(* CODESYS project Servo_Test.project

Project tree, tasks and I/O mapping:
  Device : CODESYS Virtual Control for Linux SL, CODESYS, order no. 2302000005, version 4.22.0.0
    application Application
      libraries: Standard, 3.5.22.0 (System); VisuDialogs, * (System); Unit Conversion Interfaces, * (Intern); CAA Mathematics, * (CAA Technical Workgroup); SM3_Math, * (CODESYS); SysProcess, * (System); CmpBitmapPool, * (System); SysProcess Implementation, * (System)
      task MainTask (cyclic, interval t#20ms, priority 1) calls MAIN_PRG, Ablaufkette
      task SoftMotion_PlanningTask (cyclic, interval t#2ms, priority 15) calls nothing
      global variables GVL_OPCUA
      visualisation Topics_Vis
      Structs/
        ST_RobotStatus/
          data type ST_RobotStatus
        ST_RobotAction/
          data type ST_RobotAction
          data type Error_Codes_RobotAction
        ST_RobotCommand/
          data type ST_RobotCommand
          data type Status_Codes_RobotCommand
        ST_Orientierung/
          data type ST_euler
          data type ST_quaternions
        ST_Roboter/
          data type ST_Pose_Axis
          data type ST_Pose_TCP
      old_code/
        data type Manuell_Achse
        data type TCP_Pose
        program PRG_VISU [ST]
        data type JointState
        data type ST_Servo_Axis
        data type ST_Servo_TCP
        FB_Robot/
          function block FB_Robot [FBD]
          function block FB_Watchdog [ST]
          function block FB_RobotCommander [ST]
        Interfaces/
          interface IF_RobotStatus: Ist_Pose_Axis, Ist_Pose_TCP, Ist_Mode, Client_Connection_Status, Update_Watchdog
          interface IF_RobotCommand: Soll_Pose_Axis, Soll_Pose_TCP
        function block FB_Roboter [FBD]: Update_Watchdog, Soll_Pose_Axis, Soll_Pose_TCP, Client_Connection_Status, Ist_Mode, Ist_Pose_Axis, Ist_Pose_TCP
        function block Status_POU [ST]
      program MAIN_PRG [FBD]
      FB_Generell/
        function block FB_MoveAction [ST]: MoveToHome, Ex1_ompl_tcp, Ex2_ompl_joint, Ex3_pilz_tcp_ptp, Ex_4_pilz_tcp_lin, Ablauf_HomePos, Ablauf_Pos1, Ablauf_Pos2, Ablauf_Pos3, Ablauf_Pos4, Ablauf_Pos5
        function block FB_Modes [FBD]
        function block FB_RobotStatus [ST]
        function block FB_RobotCommand [ST]
      program Ablaufkette [SFC]: Pos_6
      Funktionen/
        function FUNC_quat_to_euler [ST]
        function block FB_Quat_to_ZYZ [FBD]
        function block FB_ZYZ_to_Quat [FBD]
      Symbols
      image pool ImagePool
      visualisation VISU_Auto
      visualisation VISU_Startseite
      visualisation VISU_Manuell
      visualisation VISU_Konfig
      visualisation VISU_Schrittkette
  libraries: SM3_Robotics, * (CODESYS); VisuSymbols, 4.5.0.0 (System)
  text list GlobalTextList
*)

// Device/Application/old_code/Manuell_Achse
TYPE Manuell_Achse :
STRUCT
	axis_0_plus : BOOL;
	axis_0_minus : BOOL;
	axis_1_plus : BOOL;
	axis_1_minus : BOOL;
	axis_2_plus : BOOL;
	axis_2_minus : BOOL;
	axis_3_plus : BOOL;
	axis_3_minus : BOOL;
	axis_4_plus : BOOL;
	axis_4_minus : BOOL;
	axis_5_plus : BOOL;
	axis_5_minus : BOOL;
	//velocity_spee  einstellen
	//start manuell
END_STRUCT
END_TYPE

// Device/Application/old_code/TCP_Pose
TYPE TCP_Pose :
STRUCT
	trans_x : LREAL;
	trans_y : LREAL;
	trans_z : LREAL;
	rot_x : LREAL;
	rot_y : LREAL;
	rot_z : LREAL;
	rot_w : LREAL;
END_STRUCT
END_TYPE

//TCP Pose in kartesischen Koordinaten
//Rotation wird in quaternions uebermittelt, muss noch umgerechnet werden

// Device/Application/old_code/JointState
TYPE JointState :
STRUCT
	name :ARRAY[0..5] OF STRING;
	position :ARRAY[0..5] OF LREAL; 
	effort :ARRAY[0..5] OF LREAL;
	velocity :ARRAY[0..5] OF LREAL;
END_STRUCT
END_TYPE

// Device/Application/Structs/ST_RobotStatus/ST_RobotStatus
// Gibt den aktuellen Status des Roboters an
TYPE ST_RobotStatus :
STRUCT
	//Joints
	Ist_Pos_Axis : ST_Pose_Axis; 	
	
	// TCP mit Orientierung in Quaternions
	Ist_Pos_TCP : ST_Pose_TCP;	
	
	//Watchdog
	client_connected : BOOL;
	watchdog_counter : INT;		// Überprüft serverseitige client verbindung
END_STRUCT
END_TYPE

// Device/Application/Structs/ST_RobotCommand/ST_RobotCommand
TYPE ST_RobotCommand :
STRUCT
	// Achsen manuell verfahren
	Mode_Axis: BOOL;
	Soll_Axis_Servo : ST_Pose_Axis;
	Soll_Axis_Velocity: LREAL;
	
	// TCP manuell verfahren (funktioniert nicht, da Singularitäten auftreten wenn MoveIt Servo verwendet! Nicht in Code implementiert!)
	Mode_TCP: BOOL;
	Soll_TCP_Servo : ST_Pose_TCP;	// Hinweis: Rotation wird nur mit x,y,z übergeben und nicht als Quaternion!
	Soll_TCP_Velocity: LREAL;
	
	//enable: zum starten und stopen des services servo_node/start_servo und stop_servo
	enable : BOOL;
	
	//Status Code mit Status Codes
	Status_Code: SINT;
	
	//Watchdog
	client_connected: BOOL;
	watchdog_counter: INT;
END_STRUCT
END_TYPE

// Device/Application/Structs/ST_RobotAction/ST_RobotAction
TYPE ST_RobotAction :
STRUCT
	//Allgemein
	Execute : BOOL;					//Starten der Ausführung (Senden des Goals)
	Error_Code: DINT;				//Feedback ob Ausführung erfolgreich? (Error_code=1)

	//Planer Einstellen
	Motion_Type: STRING;			//string pipeline_id: ompl, pilz_ptp, pilz_lin 
	Planner_ID:STRING;				//string planner_id: pilz_industrial_motion_planner oder ompl
	Joint_Goal: BOOL;				
	TCP_GOAL: BOOL;
	num_planning_attempts : DINT;	//int32 num_planning_attempts
	allowed_planning_time: LREAL;	//float64 allowed_planning_time
	max_velocity_scaling: LREAL;		//float64 max_velocity_scaling_factor
	max_acceleration_scaling: LREAL;	//float64 max_acceleration_scaling_factor
	position_tolerance: LREAL;		//float 64 absolute_x_axis_tolerance ->für alle achsen die gleiche toleranz
	orientation_tolerance: LREAL;	//float64
	joint_tolerance : LREAL;
	
	//Joints
	Soll_Pos_Axis: ST_Pose_Axis;
	
	// TCP
	Soll_Pos_TCP: ST_Pose_TCP;

	//Watchdog
	client_connected : BOOL;
	watchdog_counter : INT;
END_STRUCT
END_TYPE

// Device/Application/Structs/ST_Roboter/ST_Pose_Axis
TYPE ST_Pose_Axis :
STRUCT
	axis_0 : LREAL;
	axis_1 : LREAL;
	axis_2 : LREAL;
	axis_3 : LREAL;
	axis_4 : LREAL;
	axis_5 : LREAL;
END_STRUCT
END_TYPE

// Device/Application/Structs/ST_Roboter/ST_Pose_TCP
TYPE ST_Pose_TCP :
STRUCT
	trans_x : LREAL;
	trans_y :  LREAL;
	trans_z : LREAL;
	rot_x : LREAL;
	rot_y : LREAL;
	rot_z : LREAL;
	rot_w : LREAL;
END_STRUCT
END_TYPE

// Device/Application/old_code/ST_Servo_Axis
TYPE ST_Servo_Axis :
STRUCT
	velocity : LREAL;	
	axis_0 : LREAL;
	axis_1 : LREAL;
	axis_2 : LREAL;
	axis_3 : LREAL;
	axis_4 : LREAL;
	axis_5 : LREAL;
END_STRUCT
END_TYPE

// Device/Application/old_code/ST_Servo_TCP
TYPE ST_Servo_TCP :
STRUCT
	velocity : LREAL;
	trans_x : LREAL;
	trans_y : LREAL;
	trans_z : LREAL;
	rot_x : LREAL;
	rot_y : LREAL;
	rot_z : LREAL;
	rot_w : LREAL;
END_STRUCT
END_TYPE

// Device/Application/Structs/ST_RobotAction/Error_Codes_RobotAction
{attribute 'qualified_only'}
//{attribute 'strict'}	//CODESYS erlaubt keine TYP Umwandlungen wenn strict aktiv!
{attribute 'to_string'}

TYPE Error_Codes_RobotAction :
(
	NOT_DEFINED := 0,
    SUCCESS := 1,
    FAILURE := 99999,
    PLANNING_FAILED := -1,
    INVALID_MOTION_PLAN := -2,
    MOTION_PLAN_INVALIDATED_BY_ENVIRONMENT_CHANGE := -3,
    CONTROL_FAILED := -4,
    UNABLE_TO_AQUIRE_SENSOR_DATA := -5,
    TIMED_OUT := -6,
    PREEMPTED := -7,
    START_STATE_IN_COLLISION := -10,
    START_STATE_VIOLATES_PATH_CONSTRAINTS := -11,
    START_STATE_INVALID := -26,
    GOAL_IN_COLLISION := -12,
    GOAL_VIOLATES_PATH_CONSTRAINTS := -13,
    GOAL_CONSTRAINTS_VIOLATED := -14,
    GOAL_STATE_INVALID := -27,
    UNRECOGNIZED_GOAL_TYPE := -28,
    INVALID_GROUP_NAME := -15,
    INVALID_GOAL_CONSTRAINTS := -16,
    INVALID_ROBOT_STATE := -17,
    INVALID_LINK_NAME := -18,
    INVALID_OBJECT_NAME := -19,
    FRAME_TRANSFORM_FAILURE := -21,
    COLLISION_CHECKING_UNAVAILABLE := -22,
    ROBOT_STATE_STALE := -23,
    SENSOR_INFO_STALE := -24,
    COMMUNICATION_FAILURE := -25,
    CRASH := -29,
    ABORT := -30,
    NO_IK_SOLUTION := -31
) DINT := NOT_DEFINED;	//Standardwert
END_TYPE

// Device/Application/Structs/ST_Orientierung/ST_euler
//Eulerwinkel intrinsich ZYZ
//ZYZ intrinsisch: bezug auf mitbewegendes Koordinatensystem
//ZYZ extrinsisch: bezug auf festes Koordinatensystem
TYPE ST_euler :
STRUCT
	A : LREAL;	//Z	
	B : LREAL;	//Y
	C : LREAL;	//Z
END_STRUCT
END_TYPE

// Device/Application/Structs/ST_Orientierung/ST_quaternions
TYPE ST_quaternions :
STRUCT
	qx: LREAL;
	qy: LREAL;
	qz: LREAL;
	qw: LREAL;
END_STRUCT
END_TYPE

// Device/Application/Structs/ST_RobotCommand/Status_Codes_RobotCommand
{attribute 'qualified_only'}
//{attribute 'strict'}	//CODESYS erlaubt keine TYP Umwandlungen wenn strict aktiv!
{attribute 'to_string'}
TYPE Status_Codes_RobotCommand :
(
	SERVO_AUS := 99, //wenn Roboter nicht verbunden
	INVALID := -1,
	NO_WARNING := 0,
	DECELERATE_FOR_APPROACHING_SINGULARITY := 1,
	HALT_FOR_SINGULARITY := 2,
	DECELERATE_FOR_LEAVING_SINGULARITY := 3,
	DECELERATE_FOR_COLLISION := 4,
	HALT_FOR_COLLISION := 5,
	JOINT_BOUND := 6	// Achse hat Limit erreich
) SINT := SERVO_AUS;	//Standardwert
END_TYPE

// Device/Application/GVL_OPCUA
{attribute 'qualified_only'}
VAR_GLOBAL
	//Simulation Arm
	RobotAction: ST_RobotAction;
	RobotStatus : ST_RobotStatus;
	RobotCommand : ST_RobotCommand;
	Execute : BOOL := FALSE;	//Ausführen des MoveIt2 Befehls (Auto)
	
	// Ablaufkette
	TIPP : BOOL; 				// Zum Weiterschalten
	Start_Ablaufkette: BOOL;	// Startet Ablaufkette
	Reset_Ablaufkette: BOOL;	//setzt Schrittkette zurück
	
	//Moveaction 
	Ablauf_HomePos: BOOL;
	Ablauf_Pos1: BOOL;
	Ablauf_Pos2: BOOL;
	Ablauf_Pos3: BOOL;
	Ablauf_Pos4: BOOL;
	Ablauf_Pos5: BOOL;
	
	Joint_Goal : LREAL;
	TCP_GOAL: LREAL;
	trans_x : LREAL;
	trans_y : LREAL;
	trans_z : LREAL;
	rot_A : LREAL;	
	rot_B: LREAL;
	rot_C: LREAL;	
	position_tolerance : LREAL;
	orientation_tolerance : LREAL;

	Motion_Type : STRING;
	Planner_ID : STRING;

	num_planning_attempts : LREAL;
	allowed_planning_time : LREAL;
	max_velocity_scaling : LREAL;
	max_acceleration_scaling : LREAL;



	
	//Start und Stop per "SoftKeys"
	//Übernimmt ros2 launch ... im docker container
	Start_RViz2 : BOOL;			//Start RViz2
	Stop_RViz2: BOOL;			//Stop RViz2
	Start_OPCClients: BOOL;		//Start OPC Clients
	Stop_OPC_Clients: BOOL;		//Stop OPC Clients
	

END_VAR

VAR_GLOBAL CONSTANT
	PI : REAL := 3.14159;
END_VAR

// Device/Application/MAIN_PRG
PROGRAM MAIN_PRG
VAR
///////////////////////////////////////////////////		

	//Objekt RobotAction
	RobotAction: FB_MoveAction;
	// Actions "initialisieren"
	xMoveHome : BOOL;
	xEx1_ompl_tcp: BOOL;
	xEx2_ompl_joint: BOOL;
	xEx3_pilz_tcp_ptp: BOOL;
	xEx4_pilz_tcp_lin: BOOL;
	
	//Execute trigger
	trig: R_TRIG;

	// ENUM für Error Codes
	Status_Error_Codes_Action : Error_Codes_RobotAction;
	
	Action_zyz_to_quat: FB_ZYZ_to_Quat;
///////////////////////////////////////////////////	
	
	//Modes Auswahl zur Auswahl zwischen Manuellem Modus und Automatik Modus
	Modes: FB_Modes;
	
///////////////////////////////////////////////////		

	// ObjektRobotStatus zum Anzeigen der IST Werte von Achsen und TCP
	RobotStatus: FB_RobotStatus;
	// euler : ST_Euler; für eigens programmierte Funktion
	Status_Quat_to_ZYZ: FB_Quat_to_ZYZ;
	Status_ZYZ_to_Quat : FB_ZYZ_to_Quat;
	// Status Command
	Status_Servo: Status_Codes_RobotCommand;
	
///////////////////////////////////////////////////	

	//ObjektRobotCommand zum Steuern des Roboters via MoveItServo
	// Achsen werden mit 0, 1, oder .1 angesteuert und mit velocity multipliziert
	RobotCommand: FB_RobotCommand;

END_VAR

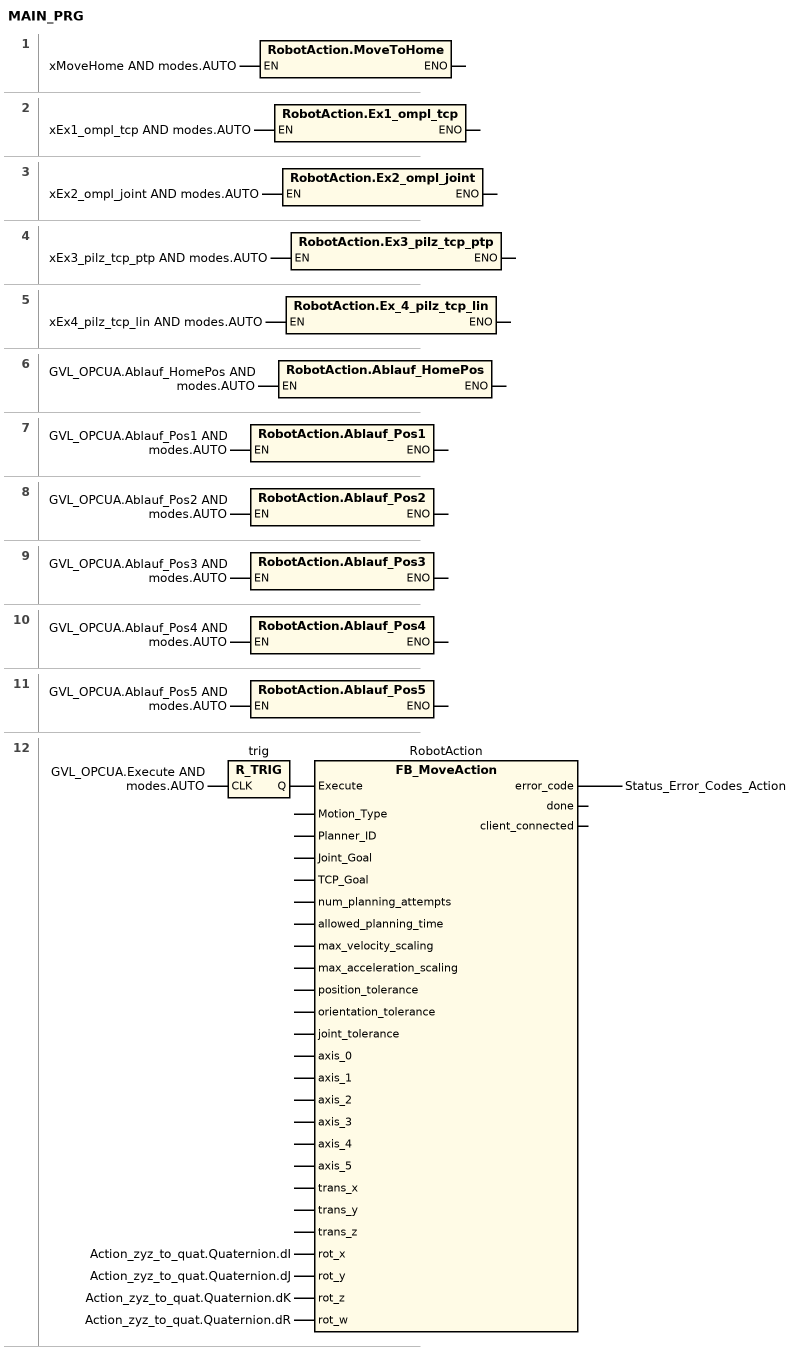
// NETWORK 1
IF xMoveHome AND modes.AUTO THEN RobotAction.MoveToHome(); END_IF

// NETWORK 2
IF xEx1_ompl_tcp AND modes.AUTO THEN RobotAction.Ex1_ompl_tcp(); END_IF

// NETWORK 3
IF xEx2_ompl_joint AND modes.AUTO THEN RobotAction.Ex2_ompl_joint(); END_IF

// NETWORK 4
IF xEx3_pilz_tcp_ptp AND modes.AUTO THEN RobotAction.Ex3_pilz_tcp_ptp(); END_IF

// NETWORK 5
IF xEx4_pilz_tcp_lin AND modes.AUTO THEN RobotAction.Ex_4_pilz_tcp_lin(); END_IF

// NETWORK 6
IF GVL_OPCUA.Ablauf_HomePos AND modes.AUTO THEN RobotAction.Ablauf_HomePos(); END_IF

// NETWORK 7
IF GVL_OPCUA.Ablauf_Pos1 AND modes.AUTO THEN RobotAction.Ablauf_Pos1(); END_IF

// NETWORK 8
IF GVL_OPCUA.Ablauf_Pos2 AND modes.AUTO THEN RobotAction.Ablauf_Pos2(); END_IF

// NETWORK 9
IF GVL_OPCUA.Ablauf_Pos3 AND modes.AUTO THEN RobotAction.Ablauf_Pos3(); END_IF

// NETWORK 10
IF GVL_OPCUA.Ablauf_Pos4 AND modes.AUTO THEN RobotAction.Ablauf_Pos4(); END_IF

// NETWORK 11
IF GVL_OPCUA.Ablauf_Pos5 AND modes.AUTO THEN RobotAction.Ablauf_Pos5(); END_IF

// NETWORK 12
trig(CLK := GVL_OPCUA.Execute AND modes.AUTO); // R_TRIG
RobotAction(
    Execute := trig.Q,
    rot_x := Action_zyz_to_quat.Quaternion.dI,
    rot_y := Action_zyz_to_quat.Quaternion.dJ,
    rot_z := Action_zyz_to_quat.Quaternion.dK,
    rot_w := Action_zyz_to_quat.Quaternion.dR); // FB_MoveAction
Status_Error_Codes_Action := RobotAction.error_code;

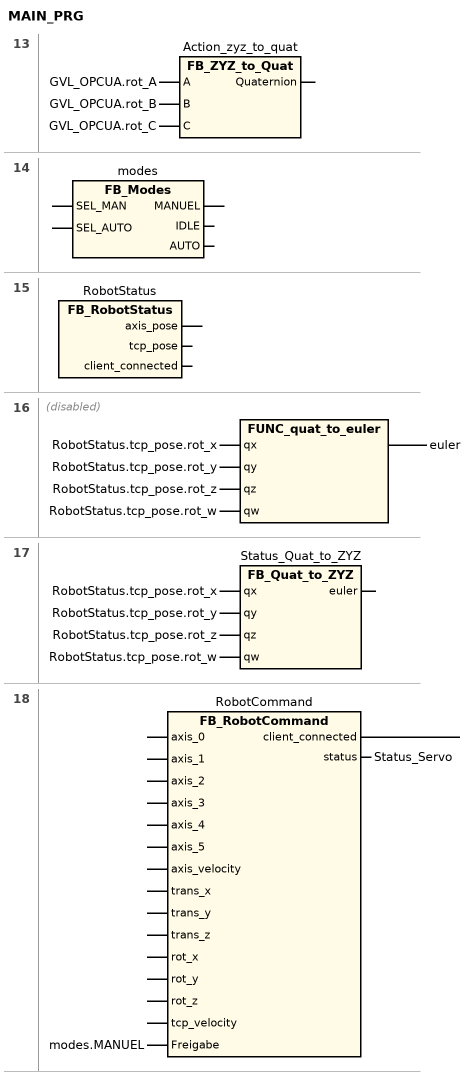
// NETWORK 13
Action_zyz_to_quat(A := GVL_OPCUA.rot_A, B := GVL_OPCUA.rot_B, C := GVL_OPCUA.rot_C); // FB_ZYZ_to_Quat

// NETWORK 14
modes(); // FB_Modes

// NETWORK 15
RobotStatus(); // FB_RobotStatus

// NETWORK 16 (disabled)
// euler := FUNC_quat_to_euler(qx := RobotStatus.tcp_pose.rot_x, qy := RobotStatus.tcp_pose.rot_y, qz := RobotStatus.tcp_pose.rot_z, qw := RobotStatus.tcp_pose.rot_w);

// NETWORK 17
Status_Quat_to_ZYZ(
    qx := RobotStatus.tcp_pose.rot_x,
    qy := RobotStatus.tcp_pose.rot_y,
    qz := RobotStatus.tcp_pose.rot_z,
    qw := RobotStatus.tcp_pose.rot_w); // FB_Quat_to_ZYZ

// NETWORK 18
RobotCommand(Freigabe := modes.MANUEL, status => Status_Servo); // FB_RobotCommand

END_PROGRAM

// Device/Application/FB_Generell/FB_MoveAction
FUNCTION_BLOCK FB_MoveAction
VAR_INPUT
    Execute : BOOL;

    Motion_Type : STRING;
    Planner_ID : STRING;

    Joint_Goal : BOOL;
    TCP_Goal : BOOL;

    num_planning_attempts : DINT;
    allowed_planning_time : LREAL;

    max_velocity_scaling : LREAL;
    max_acceleration_scaling : LREAL;

    position_tolerance : LREAL;
    orientation_tolerance : LREAL;
	joint_tolerance: LREAL;

    // Joints
    axis_0 : LREAL;
    axis_1 : LREAL;
    axis_2 : LREAL;
    axis_3 : LREAL;
    axis_4 : LREAL;
    axis_5 : LREAL;

    // TCP
    trans_x : LREAL;
    trans_y : LREAL;
    trans_z : LREAL;
    rot_x : LREAL;
    rot_y : LREAL;
    rot_z : LREAL;
    rot_w : LREAL;
	
END_VAR
VAR_OUTPUT
	error_code:DINT;
	done : BOOL;
	//Watchdog
	client_connected : BOOL;
END_VAR
VAR
	//Watchdog
	Watchdog_counter : INT;	
	Watchdog_var_old : INT := -1;
	Intervall : TIME :=T#200MS;
	Timer : TON;
	
	//Konvertierung ZYZ->Quat für action
	zyz_to_quat : FB_ZYZ_to_Quat;

END_VAR

// Execute
GVL_OPCUA.RobotAction.Execute := Execute;

// Allgemein
GVL_OPCUA.RobotAction.Motion_Type := Motion_Type;
GVL_OPCUA.RobotAction.Planner_ID := Planner_ID;

GVL_OPCUA.RobotAction.Joint_Goal := Joint_Goal;
GVL_OPCUA.RobotAction.TCP_GOAL := TCP_Goal;

GVL_OPCUA.RobotAction.num_planning_attempts := num_planning_attempts;
GVL_OPCUA.RobotAction.allowed_planning_time := allowed_planning_time;

GVL_OPCUA.RobotAction.max_velocity_scaling := max_velocity_scaling;
GVL_OPCUA.RobotAction.max_acceleration_scaling := max_acceleration_scaling;

GVL_OPCUA.RobotAction.position_tolerance := position_tolerance;
GVL_OPCUA.RobotAction.orientation_tolerance := orientation_tolerance;
GVL_OPCUA.RobotAction.joint_tolerance := joint_tolerance;

// Joints
GVL_OPCUA.RobotAction.Soll_Pos_Axis.axis_0 := axis_0;
GVL_OPCUA.RobotAction.Soll_Pos_Axis.axis_1 := axis_1;
GVL_OPCUA.RobotAction.Soll_Pos_Axis.axis_2 := axis_2;
GVL_OPCUA.RobotAction.Soll_Pos_Axis.axis_3 := axis_3;
GVL_OPCUA.RobotAction.Soll_Pos_Axis.axis_4 := axis_4;
GVL_OPCUA.RobotAction.Soll_Pos_Axis.axis_5 := axis_5;


// TCP
GVL_OPCUA.RobotAction.Soll_Pos_TCP.trans_x := trans_x;
GVL_OPCUA.RobotAction.Soll_Pos_TCP.trans_y := trans_y;
GVL_OPCUA.RobotAction.Soll_Pos_TCP.trans_z := trans_z;

GVL_OPCUA.RobotAction.Soll_Pos_TCP.rot_x := rot_x;
GVL_OPCUA.RobotAction.Soll_Pos_TCP.rot_y := rot_y;
GVL_OPCUA.RobotAction.Soll_Pos_TCP.rot_z := rot_z;
GVL_OPCUA.RobotAction.Soll_Pos_TCP.rot_w := rot_w;

//OUTPUT
error_code := GVL_OPCUA.RobotAction.Error_Code;
IF error_code = 1 THEN
	done := TRUE;
ELSE 
	done := FALSE;
END_IF

//Watchdog
Watchdog_counter := GVL_OPCUA.RobotAction.watchdog_counter;
IF Watchdog_counter <> Watchdog_var_old THEN
	Watchdog_var_old := Watchdog_counter;
	client_connected := TRUE;
	GVL_OPCUA.RobotAction.client_connected := client_connected;
	Timer(IN:=FALSE);

ELSE
	Timer(IN:=TRUE, PT:=Intervall);	
END_IF

IF Timer.Q THEN
	client_connected := FALSE;
	GVL_OPCUA.RobotAction.client_connected := client_connected;
END_IF

ACTION MoveToHome:
//HomePosition
axis_0 := 0.0;
axis_1 := 0.0;
axis_2 := 0.0;
axis_3 := 0.0;
axis_4 := 0.0;
axis_5 := 0.0;
Motion_Type := 'ompl';
Planner_ID := '';
Joint_Goal := TRUE;
TCP_Goal := FALSE;
num_planning_attempts := 5;
allowed_planning_time := 5;
max_velocity_scaling := 0.1;
max_acceleration_scaling := 0.1;
joint_tolerance := 0.005;
END_ACTION

ACTION Ex1_ompl_tcp:
trans_x := 0.114;
trans_y := -0.019;
trans_z := 0.357;
GVL_OPCUA.rot_A := 0.0;
GVL_OPCUA.rot_B := 90.0;
GVL_OPCUA.rot_C := -90.0;
Motion_Type := 'ompl';
Planner_ID := '';
Joint_Goal := FALSE;
TCP_Goal := TRUE;
num_planning_attempts := 5;
allowed_planning_time := 5;
max_velocity_scaling := 0.2;
max_acceleration_scaling := 0.2;
position_tolerance := 0.02;
orientation_tolerance := 0.05;
END_ACTION

ACTION Ex2_ompl_joint:
axis_0 := 0.1;
axis_1 := -1.65;
axis_2 := 1.7;
axis_3 := 0.1;
axis_4 := 0.2;
axis_5 := 0.3;
Motion_Type := 'ompl';
Planner_ID := '';
Joint_Goal := TRUE;
TCP_Goal := FALSE;
num_planning_attempts := 5;
allowed_planning_time := 5;
max_velocity_scaling := 0.2;
max_acceleration_scaling := 0.2;
joint_tolerance := 0.01;
END_ACTION

ACTION Ex3_pilz_tcp_ptp:
trans_x := 0.17;
trans_y := -0.04;
trans_z := 0.22;
GVL_OPCUA.rot_A := 0.0;
GVL_OPCUA.rot_B := 90.0;
GVL_OPCUA.rot_C := -90.0;
Motion_Type := 'pilz_industrial_motion_planner';
Planner_ID := 'PTP';
Joint_Goal := FALSE;
TCP_Goal := TRUE;
num_planning_attempts := 10;
allowed_planning_time := 10;
max_velocity_scaling := 0.05;
max_acceleration_scaling := 0.05;
position_tolerance := 0.02;
orientation_tolerance := 0.05;
END_ACTION

ACTION Ex_4_pilz_tcp_lin:
trans_x := 0.2;
trans_y := -0.041;
trans_z := 0.3;
GVL_OPCUA.rot_A := 0.0;
GVL_OPCUA.rot_B := 90.0;
GVL_OPCUA.rot_C := -90.0;
Motion_Type := 'pilz_industrial_motion_planner';
Planner_ID := 'LIN';
Joint_Goal := FALSE;
TCP_Goal := TRUE;
num_planning_attempts := 10;
allowed_planning_time := 10;
max_velocity_scaling := 0.005;
max_acceleration_scaling := 0.005;
position_tolerance := 0.02;
orientation_tolerance := 0.05;
END_ACTION

ACTION Ablauf_HomePos:
Joint_Goal := TRUE;
TCP_Goal := FALSE;

axis_0 := 0.1076;
axis_1 := -0.0931;
axis_2 := -1.667;
axis_3 := 1.773;
axis_4 := 0.07;
axis_5 := 0.19;

joint_tolerance := 0.01;

Motion_Type := 'ompl';
Planner_ID := '';

num_planning_attempts := 10;
allowed_planning_time := 10;

max_velocity_scaling := 0.2;
max_acceleration_scaling := 0.2;
END_ACTION

ACTION Ablauf_Pos1:
Joint_Goal := FALSE;
TCP_Goal := TRUE;

trans_x := 0.18;
trans_y := -0.0;
trans_z := 0.3;

GVL_OPCUA.rot_A := 0.0;
GVL_OPCUA.rot_B := 90.0;
GVL_OPCUA.rot_C := -90.0;

position_tolerance := 0.005;
orientation_tolerance := 0.05;

Motion_Type := 'ompl';
Planner_ID := '';

num_planning_attempts := 10;
allowed_planning_time := 10;
max_velocity_scaling := 0.1;
max_acceleration_scaling := 0.1;
END_ACTION

ACTION Ablauf_Pos2:
Joint_Goal := FALSE;
TCP_Goal := TRUE;

trans_x := 0.18;
trans_y := 0.05;
trans_z := 0.3;

GVL_OPCUA.rot_A := 0.0;
GVL_OPCUA.rot_B := 90.0;
GVL_OPCUA.rot_C := -90.0;

position_tolerance := 0.005;
orientation_tolerance := 0.05;

Motion_Type := 'pilz_industrial_motion_planner';
Planner_ID := 'PTP';


num_planning_attempts := 10;
allowed_planning_time := 10;
max_velocity_scaling := 0.1;
max_acceleration_scaling := 0.1;
END_ACTION

ACTION Ablauf_Pos3:
Joint_Goal := FALSE;
TCP_Goal := TRUE;

trans_x := 0.18;
trans_y := 0.05;
trans_z := 0.2;

GVL_OPCUA.rot_A := 0.0;
GVL_OPCUA.rot_B := 90.0;
GVL_OPCUA.rot_C := -90.0;

position_tolerance := 0.005;
orientation_tolerance := 0.05;

Motion_Type := 'pilz_industrial_motion_planner';
Planner_ID := 'PTP';


num_planning_attempts := 10;
allowed_planning_time := 10;
max_velocity_scaling := 0.1;
max_acceleration_scaling := 0.1;
END_ACTION

ACTION Ablauf_Pos4:
Joint_Goal := FALSE;
TCP_Goal := TRUE;

trans_x := 0.18;
trans_y := -0.05;
trans_z := 0.2;

GVL_OPCUA.rot_A := 0.0;
GVL_OPCUA.rot_B := 90.0;
GVL_OPCUA.rot_C := -90.0;

position_tolerance := 0.005;
orientation_tolerance := 0.05;

Motion_Type := 'pilz_industrial_motion_planner';
Planner_ID := 'PTP';


num_planning_attempts := 10;
allowed_planning_time := 10;
max_velocity_scaling := 0.1;
max_acceleration_scaling := 0.1;
END_ACTION

ACTION Ablauf_Pos5:
Joint_Goal := FALSE;
TCP_Goal := TRUE;

trans_x := 0.18;
trans_y := -0.05;
trans_z := 0.3;

GVL_OPCUA.rot_A := 0.0;
GVL_OPCUA.rot_B := 90.0;
GVL_OPCUA.rot_C := -90.0;

position_tolerance := 0.005;
orientation_tolerance := 0.05;

Motion_Type := 'pilz_industrial_motion_planner';
Planner_ID := 'PTP';


num_planning_attempts := 10;
allowed_planning_time := 10;
max_velocity_scaling := 0.1;
max_acceleration_scaling := 0.1;
END_ACTION

END_FUNCTION_BLOCK

// Device/Application/Funktionen/FB_ZYZ_to_Quat
FUNCTION_BLOCK FB_ZYZ_to_Quat
VAR_INPUT
	A : LREAL;
	B: LREAL;
	C: LREAL;
END_VAR
VAR_OUTPUT
	Quaternion: SMC_Quat;
END_VAR
VAR
	Rotation_Matrix: SMC_Matrix3;
END_VAR

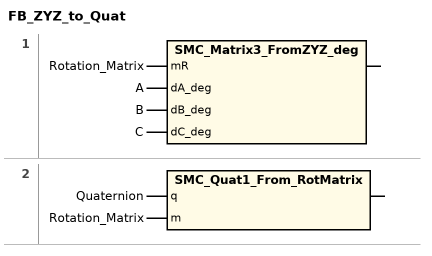
// NETWORK 1
SMC_Matrix3_FromZYZ_deg(mR := Rotation_Matrix, dA_deg := A, dB_deg := B, dC_deg := C);

// NETWORK 2
SMC_Quat1_From_RotMatrix(q := Quaternion, m := Rotation_Matrix);

END_FUNCTION_BLOCK

// Device/Application/FB_Generell/FB_Modes
FUNCTION_BLOCK FB_Modes	//mit Betriebsartenhierachie MAN > AUTO
VAR_INPUT
	SEL_MAN : BOOL;
	SEL_AUTO: BOOL;
END_VAR
VAR_OUTPUT
	MANUEL : BOOL;	//z1
	IDLE: BOOL;		//z0
	AUTO: BOOL;		//z2
END_VAR
VAR
	z0, z1, z2 : BOOL;
	H1, H2: RS;
	z: INT;
END_VAR
VAR // added by the converter: edge detectors and wires of the graphical bodies
    _w1, _w2, _w3 : BOOL;
END_VAR

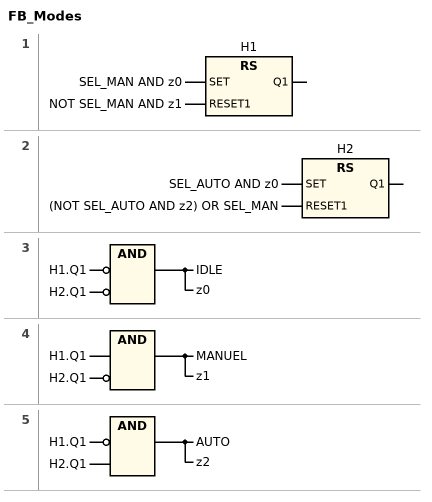
// NETWORK 1
H1(SET := SEL_MAN AND z0, RESET1 := NOT SEL_MAN AND z1); // RS

// NETWORK 2
H2(SET := SEL_AUTO AND z0, RESET1 := (NOT SEL_AUTO AND z2) OR SEL_MAN); // RS

// NETWORK 3
_w1 := NOT H1.Q1 AND NOT H2.Q1;
IDLE := _w1;
z0 := _w1;

// NETWORK 4
_w2 := H1.Q1 AND NOT H2.Q1;
MANUEL := _w2;
z1 := _w2;

// NETWORK 5
_w3 := NOT H1.Q1 AND H2.Q1;
AUTO := _w3;
z2 := _w3;

END_FUNCTION_BLOCK

// Device/Application/FB_Generell/FB_RobotStatus
FUNCTION_BLOCK FB_RobotStatus
VAR_INPUT
END_VAR
VAR_OUTPUT
	// Axis pose in RAD
	axis_pose : ST_Pose_Axis;
	
	//TCP Pose mit Orientierung in Quaternions
	tcp_pose : ST_Pose_TCP;
	
	// Watchdog
	client_connected : BOOL;
END_VAR
VAR
	//Watchdog
	Watchdog_counter : INT;	
	Watchdog_var_old : INT := -1;
	Intervall : TIME :=T#200MS;
	Timer : TON;
END_VAR

// Mappping der Variablen der GVL_OPCUA
axis_pose.axis_0 := GVL_OPCUA.RobotStatus.Ist_Pos_Axis.axis_0;
axis_pose.axis_1 := GVL_OPCUA.RobotStatus.Ist_Pos_Axis.axis_1;
axis_pose.axis_2 := GVL_OPCUA.RobotStatus.Ist_Pos_Axis.axis_2;
axis_pose.axis_3 := GVL_OPCUA.RobotStatus.Ist_Pos_Axis.axis_3;
axis_pose.axis_4 := GVL_OPCUA.RobotStatus.Ist_Pos_Axis.axis_4;
axis_pose.axis_5 := GVL_OPCUA.RobotStatus.Ist_Pos_Axis.axis_5;

tcp_pose.trans_x := GVL_OPCUA.RobotStatus.Ist_Pos_TCP.trans_x;
tcp_pose.trans_y := GVL_OPCUA.RobotStatus.Ist_Pos_TCP.trans_y;
tcp_pose.trans_z := GVL_OPCUA.RobotStatus.Ist_Pos_TCP.trans_z;
tcp_pose.rot_x := GVL_OPCUA.RobotStatus.Ist_Pos_TCP.rot_x;
tcp_pose.rot_y := GVL_OPCUA.RobotStatus.Ist_Pos_TCP.rot_y;
tcp_pose.rot_z := GVL_OPCUA.RobotStatus.Ist_Pos_TCP.rot_z;
tcp_pose.rot_w := GVL_OPCUA.RobotStatus.Ist_Pos_TCP.rot_w;

//Watchdog zum Testen ob noch mit StatusClient verbunden!
Watchdog_counter := GVL_OPCUA.RobotStatus.watchdog_counter;
IF Watchdog_counter <> Watchdog_var_old THEN
	Watchdog_var_old :=  Watchdog_counter;
    client_connected := TRUE;
	GVL_OPCUA.RobotStatus.client_connected := client_connected;
    Timer(IN := FALSE);

ELSE
    Timer(IN := TRUE,PT := Intervall );
END_IF;

IF Timer.Q THEN
    client_connected := FALSE;
	GVL_OPCUA.RobotStatus.client_connected := client_connected;
END_IF;

END_FUNCTION_BLOCK

// Device/Application/Funktionen/FUNC_quat_to_euler
FUNCTION FUNC_quat_to_euler : ST_euler
VAR_INPUT
	qx : LREAL;
	qy : LREAL;
	qz : LREAL;
	qw : LREAL;
END_VAR
VAR
	r11, r12, r13, r21, r22, r23, r31, r32, r33 : LREAL;
	const_epsilon : LREAL := 1.0E-6; // Toleranz für Gimbal Lock
	result : ST_euler;
	
END_VAR

//Quaternion -> Euler mit ZYZ (intrinsisch) 
//Ausgabe der Euler Winkel in Grad
//Rotationsmatrix Quaternion
r11 := 1.0 - 2.0 * (qy*qy + qz*qz);
r12 := 2.0 * (qx*qy - qz*qw);
r13 := 2.0 * (qx*qz + qy*qw);

r21 := 2.0 * (qx*qy + qz*qw);
r22 := 1.0 - 2.0 * (qx*qx + qz*qz);
r23 := 2.0 * (qy*qz - qx*qw);

r31 := 2.0 * (qx*qz - qy*qw);
r32 := 2.0 * (qy*qz + qx*qw);
r33 := 1.0 - 2.0 * (qx*qx + qy*qy);

result.B := MATH.atan2_func(SQRT(r31*r31+r32*r32),r33);

IF result.B < const_epsilon THEN
	//Gimbal Lock Nordpol
	result.A := 0.0;
	result.C := MATH.atan2_func(r21,r11);
	
ELSIF result.B > (MATH.PI - const_epsilon) THEN
	//Gimbal Lock Südpol
	result.A := 0.0;
	result.C := MATH.atan2_func(-r21,-r11);
ELSE
	//normal
	result.A := MATH.atan2_func(r23,r13);
	result.C := MATH.atan2_func(r32,-r31);
	
END_IF

result.A := result.A * (180.0/MATH.PI);
result.B := result.B * (180.0/MATH.PI);
result.C := result.C * (180.0/MATH.PI);

FUNC_quat_to_euler := result;

END_FUNCTION

// Device/Application/Funktionen/FB_Quat_to_ZYZ
FUNCTION_BLOCK FB_Quat_to_ZYZ
VAR_INPUT
	qx : LREAL;
	qy: LREAL;
	qz:LREAL;
	qw : LREAL;

END_VAR
VAR_OUTPUT
	euler : ST_euler;
END_VAR
VAR
	Quaternion: SMC_Quat;
	Rotation_Matrix: SMC_Matrix3;
END_VAR

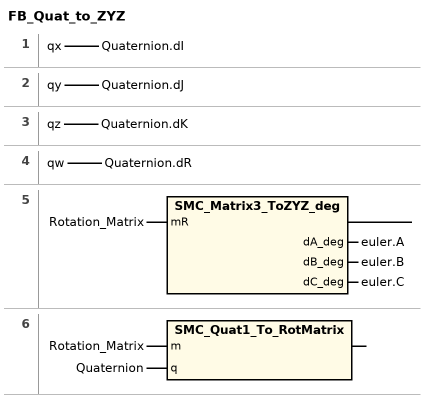
// NETWORK 1
Quaternion.dI := qx;

// NETWORK 2
Quaternion.dJ := qy;

// NETWORK 3
Quaternion.dK := qz;

// NETWORK 4
Quaternion.dR := qw;

// NETWORK 5
SMC_Matrix3_ToZYZ_deg(mR := Rotation_Matrix, dA_deg => euler.A, dB_deg => euler.B, dC_deg => euler.C);

// NETWORK 6
SMC_Quat1_To_RotMatrix(m := Rotation_Matrix, q := Quaternion);

END_FUNCTION_BLOCK

// Device/Application/FB_Generell/FB_RobotCommand
FUNCTION_BLOCK FB_RobotCommand
VAR_INPUT
	axis_0 : LREAL;
	axis_1 : LREAL;
	axis_2: LREAL;
	axis_3 : LREAL;
	axis_4 : LREAL;
	axis_5 : LREAL;
	axis_velocity : LREAL;
	
	trans_x : LREAL;
	trans_y : LREAL;
	trans_z : LREAL;
	rot_x : LREAL;
	rot_y : LREAL;
	rot_z : LREAL;
	tcp_velocity : LREAL;
	
	//Allgemein
	Freigabe:BOOL:=FALSE;
	
END_VAR
VAR_OUTPUT
	// Watchdog
	client_connected : BOOL;
	// Status Meldung
	status: SINT;	//Datentyp INT8
END_VAR
VAR
	//Watchdog
	Watchdog_counter : INT;	
	Watchdog_var_old : INT := -1;
	Intervall : TIME :=T#200MS;
	Timer : TON;
END_VAR

IF Freigabe THEN
	GVL_OPCUA.RobotCommand.Soll_Axis_Servo.axis_0 := axis_0;
	GVL_OPCUA.RobotCommand.Soll_Axis_Servo.axis_1 := axis_1;
	GVL_OPCUA.RobotCommand.Soll_Axis_Servo.axis_2 := axis_2;
	GVL_OPCUA.RobotCommand.Soll_Axis_Servo.axis_3 := axis_3;
	GVL_OPCUA.RobotCommand.Soll_Axis_Servo.axis_4 := axis_4;
	GVL_OPCUA.RobotCommand.Soll_Axis_Servo.axis_5 := axis_5;
	GVL_OPCUA.RobotCommand.Soll_Axis_Velocity := axis_velocity;
	
	GVL_OPCUA.RobotCommand.Soll_TCP_Servo.trans_x := trans_x;
	GVL_OPCUA.RobotCommand.Soll_TCP_Servo.trans_y := trans_y;
	GVL_OPCUA.RobotCommand.Soll_TCP_Servo.trans_z := trans_z;
	GVL_OPCUA.RobotCommand.Soll_TCP_Servo.rot_x := rot_x;
	GVL_OPCUA.RobotCommand.Soll_TCP_Servo.rot_y := rot_y;
	GVL_OPCUA.RobotCommand.Soll_TCP_Servo.rot_z := rot_z;
	GVL_OPCUA.RobotCommand.Soll_TCP_Velocity := tcp_velocity;
	
	// start der /servo_node/start_servo
	GVL_OPCUA.RobotCommand.enable := TRUE;
	
ELSE
	GVL_OPCUA.RobotCommand.enable := FALSE;
END_IF

// Status Code
status := GVL_OPCUA.RobotCommand.Status_Code;

//Watchdog zum Testen ob noch mit CommandClient verbunden!
Watchdog_counter := GVL_OPCUA.RobotCommand.watchdog_counter;
IF Watchdog_counter <> Watchdog_var_old THEN
	Watchdog_var_old :=  Watchdog_counter;
    client_connected := TRUE;
	GVL_OPCUA.RobotCommand.client_connected := client_connected;
    Timer(IN := FALSE);

ELSE
    Timer(IN := TRUE,PT := Intervall );
END_IF;

IF Timer.Q THEN
    client_connected := FALSE;
	GVL_OPCUA.RobotCommand.client_connected := client_connected;
END_IF;

END_FUNCTION_BLOCK

// Device/Application/Ablaufkette
PROGRAM Ablaufkette
VAR
	SFCCurrentStep : STRING;
END_VAR

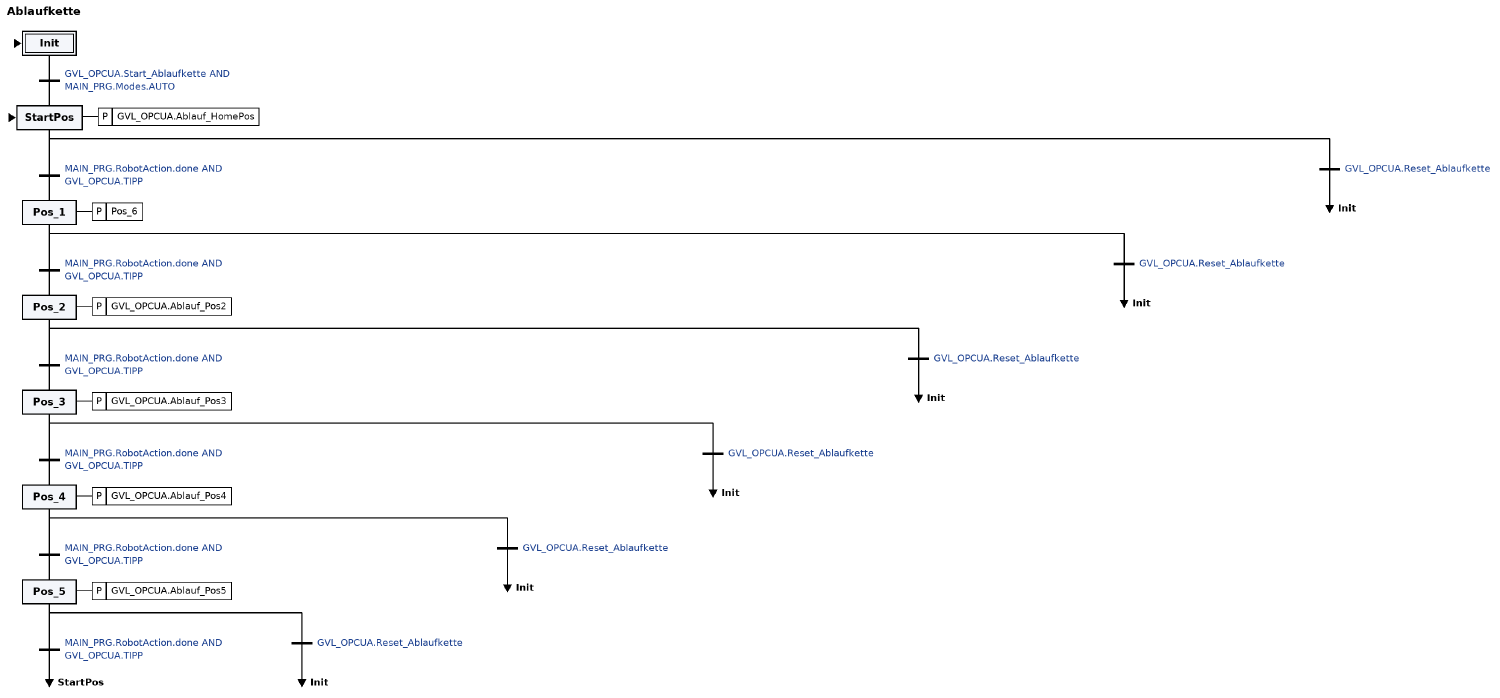
INITIAL_STEP Init:
END_STEP
TRANSITION FROM Init TO StartPos
    := GVL_OPCUA.Start_Ablaufkette AND MAIN_PRG.Modes.AUTO;
END_TRANSITION
STEP StartPos:  // min time t#1s
    GVL_OPCUA.Ablauf_HomePos(P);
END_STEP
TRANSITION FROM StartPos TO Pos_1
    := MAIN_PRG.RobotAction.done AND GVL_OPCUA.TIPP;
END_TRANSITION
TRANSITION FROM StartPos TO Init
    := GVL_OPCUA.Reset_Ablaufkette;
END_TRANSITION
STEP Pos_1:  // min time t#1s
    Pos_6(P);
END_STEP
TRANSITION FROM Pos_1 TO Pos_2
    := MAIN_PRG.RobotAction.done AND GVL_OPCUA.TIPP;
END_TRANSITION
TRANSITION FROM Pos_1 TO Init
    := GVL_OPCUA.Reset_Ablaufkette;
END_TRANSITION
STEP Pos_2:  // min time t#1s
    GVL_OPCUA.Ablauf_Pos2(P);
END_STEP
TRANSITION FROM Pos_2 TO Pos_3
    := MAIN_PRG.RobotAction.done AND GVL_OPCUA.TIPP;
END_TRANSITION
TRANSITION FROM Pos_2 TO Init
    := GVL_OPCUA.Reset_Ablaufkette;
END_TRANSITION
STEP Pos_3:  // min time t#1s
    GVL_OPCUA.Ablauf_Pos3(P);
END_STEP
TRANSITION FROM Pos_3 TO Pos_4
    := MAIN_PRG.RobotAction.done AND GVL_OPCUA.TIPP;
END_TRANSITION
TRANSITION FROM Pos_3 TO Init
    := GVL_OPCUA.Reset_Ablaufkette;
END_TRANSITION
STEP Pos_4:  // min time t#1s
    GVL_OPCUA.Ablauf_Pos4(P);
END_STEP
TRANSITION FROM Pos_4 TO Pos_5
    := MAIN_PRG.RobotAction.done AND GVL_OPCUA.TIPP;
END_TRANSITION
TRANSITION FROM Pos_4 TO Init
    := GVL_OPCUA.Reset_Ablaufkette;
END_TRANSITION
STEP Pos_5:  // min time t#1s
    GVL_OPCUA.Ablauf_Pos5(P);
END_STEP
TRANSITION FROM Pos_5 TO StartPos
    := MAIN_PRG.RobotAction.done AND GVL_OPCUA.TIPP;
END_TRANSITION
TRANSITION FROM Pos_5 TO Init
    := GVL_OPCUA.Reset_Ablaufkette;
END_TRANSITION

ACTION Pos_6:
MAIN_PRG.RobotAction.Joint_Goal := FALSE;
MAIN_PRG.RobotAction.TCP_Goal := TRUE;

MAIN_PRG.RobotAction.trans_x := 0.18;
MAIN_PRG.RobotAction.trans_y := -0.0;
MAIN_PRG.RobotAction.trans_z := 0.3;

GVL_OPCUA.rot_A := 0.0;
GVL_OPCUA.rot_B := 90.0;
GVL_OPCUA.rot_C := -90.0;

MAIN_PRG.RobotAction.position_tolerance := 0.005;
MAIN_PRG.RobotAction.orientation_tolerance := 0.05;

MAIN_PRG.RobotAction.Motion_Type := 'ompl';
MAIN_PRG.RobotAction.Planner_ID := '';

MAIN_PRG.RobotAction.num_planning_attempts := 10;
MAIN_PRG.RobotAction.allowed_planning_time := 10;
MAIN_PRG.RobotAction.max_velocity_scaling := 0.1;
MAIN_PRG.RobotAction.max_acceleration_scaling := 0.1;
END_ACTION

END_PROGRAM

// Device/Application/old_code/PRG_VISU
PROGRAM PRG_Visu
VAR
    //arrStruct: ARRAY[0..6] OF LREAL;
	Robot : FB_Robot;
	
	//Instanziierung für Roboter
	axis_0_plus :BOOL := FALSE;
	axis_0_minus :BOOL := FALSE;
	axis_1_plus :BOOL := FALSE;
	axis_1_minus :BOOL := FALSE;
	axis_2_plus :BOOL := FALSE;
	axis_2_minus :BOOL := FALSE;
	axis_3_plus :BOOL := FALSE;
	axis_3_minus :BOOL := FALSE;
	axis_4_plus :BOOL := FALSE;
	axis_4_minus :BOOL := FALSE;
	axis_5_plus :BOOL := FALSE;
	axis_5_minus :BOOL := FALSE;
	vis_velocity :LREAL := 0;
END_VAR

Robot();

END_PROGRAM

// Device/Application/old_code/FB_Robot/FB_Robot
FUNCTION_BLOCK FB_Robot
VAR_INPUT
	Command: RobotCommand;
END_VAR
VAR_OUTPUT
	Status: ST_RobotStatus;
END_VAR
VAR
	robotcommand : FB_RobotCommand;
	Watchdog: FB_Watchdog;
END_VAR

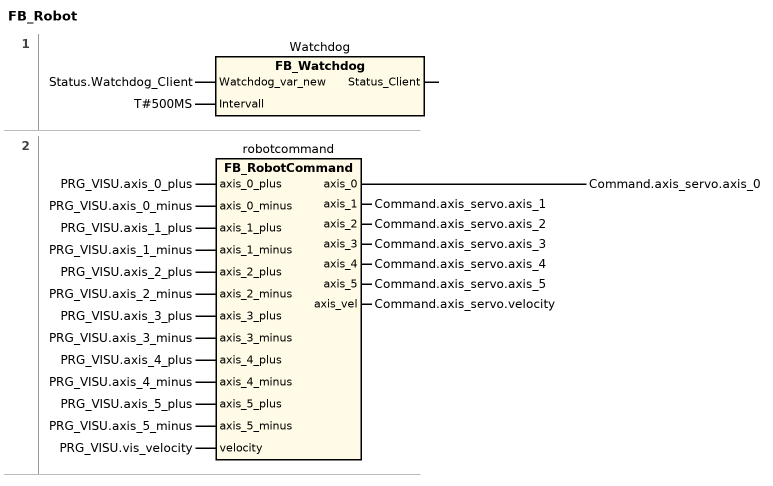
// NETWORK 1
Watchdog(Watchdog_var_new := Status.Watchdog_Client, Intervall := T#500MS); // FB_Watchdog

// NETWORK 2
robotcommand(
    axis_0_plus := PRG_VISU.axis_0_plus,
    axis_0_minus := PRG_VISU.axis_0_minus,
    axis_1_plus := PRG_VISU.axis_1_plus,
    axis_1_minus := PRG_VISU.axis_1_minus,
    axis_2_plus := PRG_VISU.axis_2_plus,
    axis_2_minus := PRG_VISU.axis_2_minus,
    axis_3_plus := PRG_VISU.axis_3_plus,
    axis_3_minus := PRG_VISU.axis_3_minus,
    axis_4_plus := PRG_VISU.axis_4_plus,
    axis_4_minus := PRG_VISU.axis_4_minus,
    axis_5_plus := PRG_VISU.axis_5_plus,
    axis_5_minus := PRG_VISU.axis_5_minus,
    velocity := PRG_VISU.vis_velocity,
    axis_1 => Command.axis_servo.axis_1,
    axis_2 => Command.axis_servo.axis_2,
    axis_3 => Command.axis_servo.axis_3,
    axis_4 => Command.axis_servo.axis_4,
    axis_5 => Command.axis_servo.axis_5,
    axis_vel => Command.axis_servo.velocity); // FB_RobotCommand
Command.axis_servo.axis_0 := robotcommand.axis_0;

END_FUNCTION_BLOCK

// Device/Application/old_code/FB_Robot/FB_Watchdog
FUNCTION_BLOCK FB_Watchdog
VAR_INPUT
	Watchdog_var_new: INT;
	Intervall : TIME;
END_VAR
VAR_OUTPUT
	Status_Client : BOOL;
END_VAR
VAR
	Watchdog_var_old : INT := -1;
	Timer : TON;
END_VAR

IF Watchdog_var_new <> Watchdog_var_old THEN

    Watchdog_var_old := Watchdog_var_new;
    Status_Client := TRUE;
    Timer(IN := FALSE);

ELSE
    Timer(IN := TRUE,PT := Intervall );
END_IF;

IF Timer.Q THEN
    Status_Client := FALSE;
END_IF;

END_FUNCTION_BLOCK

// Device/Application/old_code/FB_Robot/FB_RobotCommander
FUNCTION_BLOCK FB_RobotCommander
VAR_INPUT
	axis_0_plus : BOOL;
	axis_0_minus : BOOL;
	axis_1_plus : BOOL;
	axis_1_minus : BOOL;
	axis_2_plus : BOOL;
	axis_2_minus : BOOL;
	axis_3_plus : BOOL;
	axis_3_minus : BOOL;
	axis_4_plus : BOOL;
	axis_4_minus : BOOL;
	axis_5_plus : BOOL;
	axis_5_minus : BOOL;
	velocity : LREAL;
END_VAR
VAR_OUTPUT
	axis_0 : LREAL;
	axis_1 : LREAL;
	axis_2 : LREAL;
	axis_3 : LREAL;
	axis_4 : LREAL;
	axis_5 : LREAL;
	axis_vel : LREAL;
END_VAR
VAR
END_VAR

// Achse 0
IF axis_0_plus THEN
    axis_0 := 1;
ELSIF axis_0_minus THEN
    axis_0 := -1;
ELSE
    axis_0 := 0;
END_IF;

// Achse 1
IF axis_1_plus THEN
    axis_1 := 1;
ELSIF axis_1_minus THEN
    axis_1 := -1;
ELSE
    axis_1 := 0;
END_IF;

// Achse 2
IF axis_2_plus THEN
    axis_2 := 1;
ELSIF axis_2_minus THEN
    axis_2 := -1;
ELSE
    axis_2 := 0;
END_IF;

// Achse 3
IF axis_3_plus THEN
    axis_3 := 1;
ELSIF axis_3_minus THEN
    axis_3 := -1;
ELSE
    axis_3 := 0;
END_IF;

// Achse 4
IF axis_4_plus THEN
    axis_4 := 1;
ELSIF axis_4_minus THEN
    axis_4 := -1;
ELSE
    axis_4 := 0;
END_IF;

// Achse 5
IF axis_5_plus THEN
    axis_5 := 1;
ELSIF axis_5_minus THEN
    axis_5 := -1;
ELSE
    axis_5 := 0;
END_IF;

// Geschwimdigkeit setzten
axis_vel := velocity;

END_FUNCTION_BLOCK

// Device/Application/old_code/Interfaces/IF_RobotStatus
INTERFACE IF_RobotStatus

PROPERTY Ist_Pose_Axis : ST_Pose_Axis
GET
END_GET
END_PROPERTY

PROPERTY Ist_Pose_TCP : ST_Pose_TCP
GET
END_GET
END_PROPERTY

PROPERTY Ist_Mode : ST_Modes
SET
END_SET
GET
END_GET
END_PROPERTY

PROPERTY Client_Connection_Status : BOOL
SET
END_SET
GET
END_GET
END_PROPERTY

METHOD Update_Watchdog : BOOL
VAR_INPUT
END_VAR
END_METHOD

END_INTERFACE

// Device/Application/old_code/Interfaces/IF_RobotCommand
INTERFACE IF_RobotCommand

PROPERTY Soll_Pose_Axis : ST_Servo_Axis
SET
END_SET
GET
END_GET
END_PROPERTY

PROPERTY Soll_Pose_TCP : ST_Servo_TCP
SET
END_SET
GET
END_GET
END_PROPERTY

END_INTERFACE

// Device/Application/old_code/FB_Roboter
FUNCTION_BLOCK FB_Roboter IMPLEMENTS IF_RobotCommand, IF_RobotStatus
VAR_INPUT
END_VAR
VAR_OUTPUT
END_VAR
VAR
	// --- Command Variablen ---
    _soll_pose_axis : ST_Servo_Axis; // (Passend zu deinem Struct-Namen)
    _soll_pose_tcp  : ST_Servo_TCP;
    
    // --- Status Variablen ---
    _client_connected : BOOL;
    _ist_mode         : ST_Modes;
    _ist_pose_axis    : ST_Pose_Axis;
    _ist_pose_tcp     : ST_Pose_TCP;
END_VAR

// NETWORK 1

{warning 'Methodenimplementierung hinzufügen'}
METHOD Update_Watchdog : BOOL
END_METHOD

{warning 'Eigenschaftenimplementierung hinzufügen'}
PROPERTY Soll_Pose_Axis : ST_Servo_Axis
GET
END_GET
SET
END_SET
END_PROPERTY

{warning 'Eigenschaftenimplementierung hinzufügen'}
PROPERTY Soll_Pose_TCP : ST_Servo_TCP
GET
END_GET
SET
END_SET
END_PROPERTY

{warning 'Eigenschaftenimplementierung hinzufügen'}
PROPERTY Client_Connection_Status : BOOL
GET
END_GET
SET
END_SET
END_PROPERTY

{warning 'Eigenschaftenimplementierung hinzufügen'}
PROPERTY Ist_Mode : ST_Modes
GET
END_GET
SET
END_SET
END_PROPERTY

{warning 'Eigenschaftenimplementierung hinzufügen'}
PROPERTY Ist_Pose_Axis : ST_Pose_Axis
GET
END_GET
SET
END_SET
END_PROPERTY

{warning 'Eigenschaftenimplementierung hinzufügen'}
PROPERTY Ist_Pose_TCP : ST_Pose_TCP
GET
END_GET
SET
END_SET
END_PROPERTY

END_FUNCTION_BLOCK

// Device/Application/old_code/Status_POU
FUNCTION_BLOCK Status_POU
VAR_IN_OUT
END_VAR
VAR_OUTPUT
	Status : ST_RobotStatus;
END_VAR
VAR
END_VAR

END_FUNCTION_BLOCK

// Device/Application/Topics_Vis
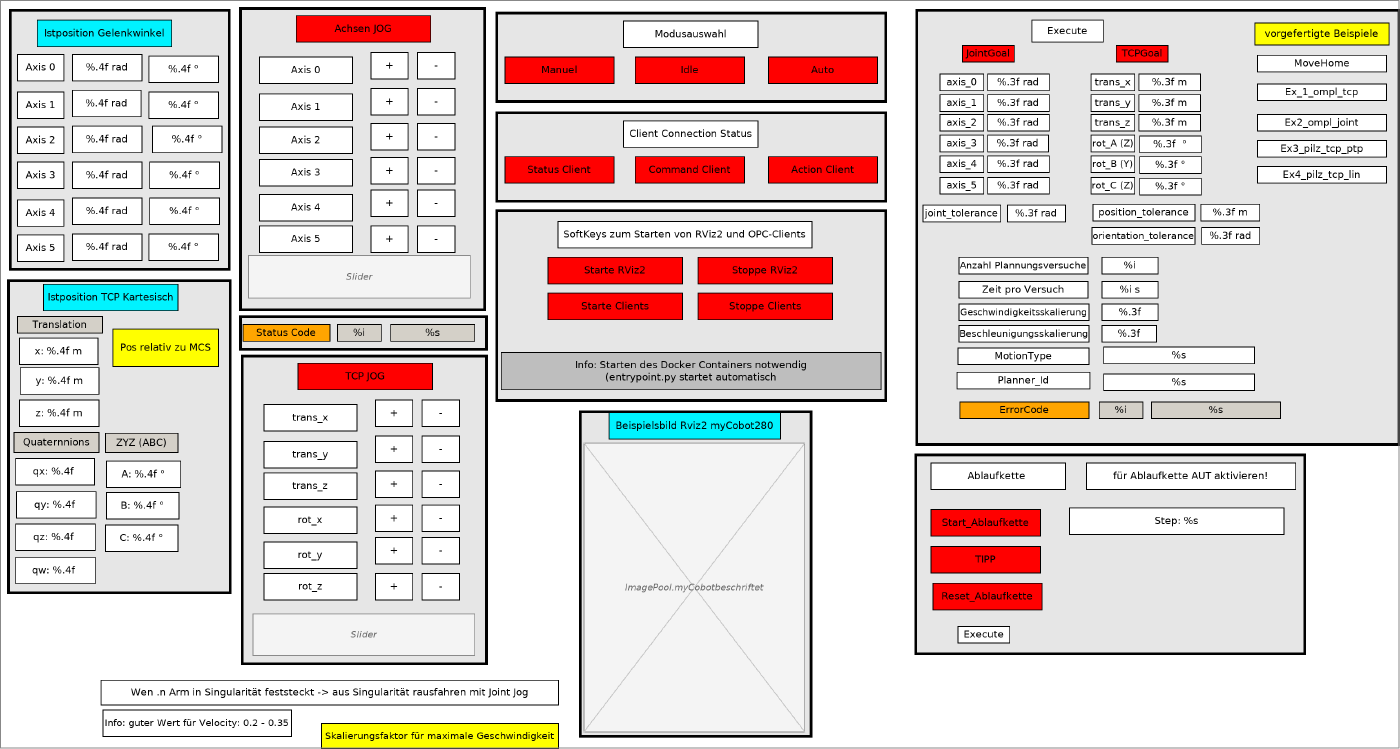
VISUALIZATION Topics_Vis  // 1557x834
    Rectangle (266,351 276x39)
    Rectangle (266,8 274x338)
    Rectangle (644,457 259x364)
    Rectangle (551,233 435x214)
    Rectangle (8,311 249x350)
    Rectangle (1018,10 539x486)
    Rectangle (551,13 435x101)
    Rectangle (10,10 246x291)
    Rectangle (41,22 150x30), "Istposition Gelenkwinkel"
    Rectangle (48,316 150x30), "Istposition TCP Kartesisch"
    Rectangle (21,376 88x30), "x: %.4f m", text variable: MAIN_PRG.RobotStatus.tcp_pose.trans_x
    Rectangle (22,409 88x30), "y: %.4f m", text variable: MAIN_PRG.RobotStatus.tcp_pose.trans_y
    Rectangle (21,445 89x30), "z: %.4f m", text variable: MAIN_PRG.RobotStatus.tcp_pose.trans_z
    Rectangle (17,510 88x30), "qx: %.4f", text variable: MAIN_PRG.RobotStatus.tcp_pose.rot_x
    Rectangle (18,547 89x30), "qy: %.4f", text variable: MAIN_PRG.RobotStatus.tcp_pose.rot_y
    Rectangle (17,583 89x30), "qz: %.4f", text variable: MAIN_PRG.RobotStatus.tcp_pose.rot_z
    Rectangle (17,620 89x30), "qw: %.4f", text variable: MAIN_PRG.RobotStatus.tcp_pose.rot_w
    Rectangle (412,58 42x30), "+"
        OnMouseDown: execute { MAIN_PRG.RobotCommand.axis_0 := +1; }
        OnMouseUp: execute { MAIN_PRG.RobotCommand.axis_0 := 0; }
    Rectangle (464,58 42x30), "-"
        OnMouseDown: execute { MAIN_PRG.RobotCommand.axis_0 := -1; }
        OnMouseUp: execute { MAIN_PRG.RobotCommand.axis_0 := 0; }
    Rectangle (412,98 42x30), "+"
        OnMouseDown: execute { MAIN_PRG.RobotCommand.axis_1 := +1; }
        OnMouseUp: execute { MAIN_PRG.RobotCommand.axis_1 := 0; }
    Rectangle (464,137 42x30), "-"
        OnMouseDown: execute { MAIN_PRG.RobotCommand.axis_2 := -1; }
        OnMouseUp: execute { MAIN_PRG.RobotCommand.axis_2 := 0; }
    Rectangle (412,137 42x30), "+"
        OnMouseDown: execute { MAIN_PRG.RobotCommand.axis_2 := +1; }
        OnMouseUp: execute { MAIN_PRG.RobotCommand.axis_2 := 0; }
    Rectangle (412,175 42x30), "+"
        OnMouseDown: execute { MAIN_PRG.RobotCommand.axis_3 := +1; }
        OnMouseUp: execute { MAIN_PRG.RobotCommand.axis_3 := 0; }
    Rectangle (464,98 42x30), "-"
        OnMouseDown: execute { MAIN_PRG.RobotCommand.axis_1 := -1; }
        OnMouseUp: execute { MAIN_PRG.RobotCommand.axis_1 := 0; }
    Rectangle (464,175 42x30), "-"
        OnMouseDown: execute { MAIN_PRG.RobotCommand.axis_3 := -1; }
        OnMouseUp: execute { MAIN_PRG.RobotCommand.axis_3 := 0; }
    Rectangle (412,211 42x30), "+"
        OnMouseDown: execute { MAIN_PRG.RobotCommand.axis_4 := +1; }
        OnMouseUp: execute { MAIN_PRG.RobotCommand.axis_4 := 0; }
    Rectangle (464,211 42x30), "-"
        OnMouseDown: execute { MAIN_PRG.RobotCommand.axis_4 := -1; }
        OnMouseUp: execute { MAIN_PRG.RobotCommand.axis_4 := 0; }
    Rectangle (412,251 42x30), "+"
        OnMouseDown: execute { MAIN_PRG.RobotCommand.axis_5 := +1; }
        OnMouseUp: execute { MAIN_PRG.RobotCommand.axis_5 := 0; }
    Rectangle (464,251 42x30), "-"
        OnMouseDown: execute { MAIN_PRG.RobotCommand.axis_5 := -1; }
        OnMouseUp: execute { MAIN_PRG.RobotCommand.axis_5 := 0; }
    Slider (276,284 247x48), variable: MAIN_PRG.RobotCommand.axis_velocity, scale 0..1
    Rectangle (693,23 150x30), "Modusauswahl"
    Rectangle (80,60 78x30), "%.4f rad", text variable: MAIN_PRG.RobotStatus.axis_pose.axis_0
    Rectangle (80,100 77x30), "%.4f rad", text variable: MAIN_PRG.RobotStatus.axis_pose.axis_1
    Rectangle (80,140 78x30), "%.4f rad", text variable: MAIN_PRG.RobotStatus.axis_pose.axis_2
    Rectangle (80,180 78x30), "%.4f rad", text variable: MAIN_PRG.RobotStatus.axis_pose.axis_3
    Rectangle (80,220 78x30), "%.4f rad", text variable: MAIN_PRG.RobotStatus.axis_pose.axis_4
    Rectangle (80,260 78x30), "%.4f rad", text variable: MAIN_PRG.RobotStatus.axis_pose.axis_5
    Rectangle (329,17 150x30), "Achsen JOG", colour toggle: GVL_OPCUA.RobotCommand.Mode_Axis
        toggle GVL_OPCUA.RobotCommand.Mode_Axis
        OnMouseClick: execute { GVL_OPCUA.RobotCommand.Mode_TCP := FALSE; }
    Rectangle (561,63 122x30), "Manuel", colour toggle: MAIN_PRG.Modes.MANUEL
        toggle MAIN_PRG.Modes.SEL_MAN p2164770859=TRUE
    Rectangle (854,63 122x30), "Auto", colour toggle: MAIN_PRG.Modes.AUTO
        toggle MAIN_PRG.Modes.SEL_AUTO p2164770859=TRUE
    Rectangle (706,63 122x30), "Idle", colour toggle: MAIN_PRG.Modes.IDLE
    Rectangle (1045,82 49x19), "axis_0"
    Rectangle (1045,105 49x19), "axis_1"
    Rectangle (1045,127 49x19), "axis_2"
    Rectangle (1045,150 49x19), "axis_3"
    Rectangle (1045,173 49x19), "axis_4"
    Rectangle (1045,197 49x19), "axis_5"
    Rectangle (1098,82 69x19), "%.3f rad", text variable: MAIN_PRG.RobotAction.axis_0
        OnMouseClick: write the text variable via Default
    Rectangle (1098,105 69x19), "%.3f rad", text variable: MAIN_PRG.RobotAction.axis_1
        OnMouseClick: write the text variable via Default
    Rectangle (1098,127 69x19), "%.3f rad", text variable: MAIN_PRG.RobotAction.axis_2
        OnMouseClick: write the text variable via Default
    Rectangle (1098,150 68x19), "%.3f rad", text variable: MAIN_PRG.RobotAction.axis_3
        OnMouseClick: write the text variable via Default
    Rectangle (1098,173 69x19), "%.3f rad", text variable: MAIN_PRG.RobotAction.axis_4
        OnMouseClick: write the text variable via Default
    Rectangle (1098,197 69x19), "%.3f rad", text variable: MAIN_PRG.RobotAction.axis_5
        OnMouseClick: write the text variable via Default
    Rectangle (1213,82 49x19), "trans_x"
    Rectangle (1213,105 49x19), "trans_y"
    Rectangle (1213,127 49x19), "trans_z"
    Rectangle (1266,82 69x19), "%.3f m", text variable: MAIN_PRG.RobotAction.trans_x
        OnMouseClick: write the text variable via Default
    Rectangle (1266,105 69x19), "%.3f m", text variable: MAIN_PRG.RobotAction.trans_y
        OnMouseClick: write the text variable via Default
    Rectangle (1266,127 69x19), "%.3f m", text variable: MAIN_PRG.RobotAction.trans_z
        OnMouseClick: write the text variable via Default
    Rectangle (1147,22 80x25), "Execute"
        tap GVL_OPCUA.Execute
    Rectangle (1070,50 58x19), "JointGoal", colour toggle: MAIN_PRG.RobotAction.Joint_Goal
        toggle MAIN_PRG.RobotAction.Joint_Goal
    Rectangle (1241,50 58x19), "TCPGoal", colour toggle: MAIN_PRG.RobotAction.TCP_Goal
        toggle MAIN_PRG.RobotAction.TCP_Goal
    Rectangle (1066,286 144x19), "Anzahl Plannungsversuche"
    Rectangle (1066,313 144x19), "Zeit pro Versuch"
    Rectangle (1066,338 145x19), "Geschwindigkeitsskalierung"
    Rectangle (1066,362 145x19), "Beschleunigungsskalierung"
    Rectangle (1215,227 114x19), "position_tolerance"
    Rectangle (1214,253 115x19), "orientation_tolerance"
    Rectangle (1225,286 63x19), "%i", text variable: MAIN_PRG.RobotAction.num_planning_attempts
        OnMouseClick: write the text variable via Default
    Rectangle (1225,313 63x19), "%i s", text variable: MAIN_PRG.RobotAction.allowed_planning_time
        OnMouseClick: write the text variable via Default
    Rectangle (1225,338 63x19), "%.3f", text variable: MAIN_PRG.RobotAction.max_velocity_scaling
        OnMouseClick: write the text variable via Default
    Rectangle (1225,362 61x19), "%.3f", text variable: MAIN_PRG.RobotAction.max_acceleration_scaling
        OnMouseClick: write the text variable via Default
    Rectangle (1335,227 66x19), "%.3f m", text variable: MAIN_PRG.RobotAction.position_tolerance
        OnMouseClick: write the text variable via Default
    Rectangle (1336,253 65x19), "%.3f rad", text variable: MAIN_PRG.RobotAction.orientation_tolerance
        OnMouseClick: write the text variable via Default
    Rectangle (1065,387 146x19), "MotionType"
    Rectangle (1064,414 148x19), "Planner_Id"
    Rectangle (1067,447 144x19), "ErrorCode"
    Rectangle (1222,447 49x19), "%i", text variable: MAIN_PRG.RobotAction.error_code
    Rectangle (1227,386 168x19), "%s", text variable: MAIN_PRG.RobotAction.Motion_Type
        OnMouseClick: write the text variable via Default
    Rectangle (1227,416 168x19), "%s", text variable: MAIN_PRG.RobotAction.Planner_ID
        OnMouseClick: write the text variable via Default
    Rectangle (1398,61 144x19), "MoveHome"
        tap MAIN_PRG.xMoveHome
    Rectangle (1280,447 144x19), "%s", text variable: MAIN_PRG.Status_Error_Codes_Action
    Rectangle (551,124 435x101)
    Rectangle (693,134 150x30), "Client Connection Status"
    Rectangle (561,174 122x30), "Status Client", colour toggle: MAIN_PRG.RobotStatus.client_connected
    Rectangle (854,174 122x30), "Action Client", colour toggle: MAIN_PRG.RobotAction.client_connected
    Rectangle (706,174 122x30), "Command Client", colour toggle: MAIN_PRG.RobotCommand.client_connected
    Rectangle (1398,93 144x19), "Ex_1_ompl_tcp"
        tap MAIN_PRG.xEx1_ompl_tcp
    Rectangle (1398,127 144x19), "Ex2_ompl_joint"
        tap MAIN_PRG.xEx2_ompl_joint
    Rectangle (1398,156 144x19), "Ex3_pilz_tcp_ptp"
        tap MAIN_PRG.xEx3_pilz_tcp_ptp
    Rectangle (1398,185 144x19), "Ex4_pilz_tcp_lin"
        tap MAIN_PRG.xEx4_pilz_tcp_lin
    Rectangle (165,62 78x30), "%.4f °", text variable: MAIN_PRG.RobotStatus.axis_pose.axis_0 *(180.0/GVL_OPCUA.PI)
    Rectangle (165,102 78x30), "%.4f °", text variable: MAIN_PRG.RobotStatus.axis_pose.axis_1 *(180.0/GVL_OPCUA.PI)
    Rectangle (169,140 78x30), "%.4f °", text variable: MAIN_PRG.RobotStatus.axis_pose.axis_2 *(180.0/GVL_OPCUA.PI)
    Rectangle (166,180 78x30), "%.4f °", text variable: MAIN_PRG.RobotStatus.axis_pose.axis_3 *(180.0/GVL_OPCUA.PI)
    Rectangle (166,220 78x30), "%.4f °", text variable: MAIN_PRG.RobotStatus.axis_pose.axis_4 *(180.0/GVL_OPCUA.PI)
    Rectangle (165,260 78x30), "%.4f °", text variable: MAIN_PRG.RobotStatus.axis_pose.axis_5 *(180.0/GVL_OPCUA.PI)
    Rectangle (118,513 83x30), "A: %.4f °", text variable: MAIN_PRG.Status_Quat_to_ZYZ.euler.A
    Rectangle (118,548 81x30), "B: %.4f °", text variable: MAIN_PRG.Status_Quat_to_ZYZ.euler.B
    Rectangle (117,584 81x30), "C: %.4f °", text variable: MAIN_PRG.Status_Quat_to_ZYZ.euler.C
    Rectangle (117,482 81x22), "ZYZ (ABC)"
    Rectangle (1017,505 435x224)
    Rectangle (1035,515 150x30), "Ablaufkette"
    Rectangle (1035,608 122x30), "TIPP", colour toggle: MAIN_PRG.RobotStatus.client_connected
        tap GVL_OPCUA.TIPP
    Rectangle (1035,567 122x30), "Start_Ablaufkette", colour toggle: MAIN_PRG.RobotStatus.client_connected
        tap GVL_OPCUA.Start_Ablaufkette
    Rectangle (1189,565 239x30), "Step: %s", text variable: Ablaufkette.SFCCurrentStep
    Rectangle (1208,515 233x30), "für Ablaufkette AUT aktivieren!"
    Rectangle (1037,649 122x30), "Reset_Ablaufkette", colour toggle: MAIN_PRG.RobotStatus.client_connected
        tap GVL_OPCUA.Reset_Ablaufkette
    Rectangle (1065,697 58x19), "Execute"
        tap GVL_OPCUA.Execute
    Rectangle (15,481 95x23), "Quaternnions"
    Rectangle (609,286 150x30), "Starte RViz2"
        toggle GVL_OPCUA.Start_RViz2
    Rectangle (609,326 150x30), "Starte Clients"
        toggle GVL_OPCUA.Start_OPCClients
    Rectangle (776,326 150x30), "Stoppe Clients"
        toggle GVL_OPCUA.Stop_OPC_Clients
    Rectangle (776,286 150x30), "Stoppe RViz2"
        toggle GVL_OPCUA.Stop_RViz2
    Rectangle (288,63 104x30), "Axis 0"
    Rectangle (288,104 104x30), "Axis 1"
    Rectangle (288,141 104x30), "Axis 2"
    Rectangle (288,177 104x30), "Axis 3"
    Rectangle (288,216 104x30), "Axis 4"
    Rectangle (288,251 104x30), "Axis 5"
    Rectangle (19,60 52x30), "Axis 0"
    Rectangle (19,102 52x30), "Axis 1"
    Rectangle (19,141 52x30), "Axis 2"
    Rectangle (19,180 52x30), "Axis 3"
    Rectangle (19,222 52x30), "Axis 4"
    Rectangle (19,261 52x30), "Axis 5"
    RoundedRectangle (125,366 118x42), "Pos relativ zu MCS"
    Image (649,493 246x322), image: ImagePool.myCobotbeschriftet
    Rectangle (677,459 191x30), "Beispielsbild Rviz2 myCobot280"
    RoundedRectangle (1395,25 150x25), "vorgefertigte Beispiele"
    Rectangle (620,246 283x30), "SoftKeys zum Starten von RViz2 und OPC-Clients"
    Rectangle (557,392 423x42), "Info: Starten des Docker Containers notwendig (entrypoint.py startet automatisch"
    Rectangle (1213,150 49x19), "rot_A (Z)"
    Rectangle (1213,173 49x19), "rot_B (Y)"
    Rectangle (1213,197 49x19), "rot_C (Z)"
    Rectangle (1267,151 69x19), "%.3f °", text variable: GVL_OPCUA.rot_A
        OnMouseClick: write the text variable via Default
    Rectangle (1267,174 69x19), "%.3f °", text variable: GVL_OPCUA.rot_B
        OnMouseClick: write the text variable via Default
    Rectangle (1267,198 69x19), "%.3f °", text variable: GVL_OPCUA.rot_C
        OnMouseClick: write the text variable via Default
    Rectangle (1026,228 87x19), "joint_tolerance"
    Rectangle (1120,228 65x19), "%.3f rad", text variable: MAIN_PRG.RobotAction.joint_tolerance
        OnMouseClick: write the text variable via Default
    Rectangle (268,395 274x345)
    Rectangle (417,445 42x30), "+"
        OnMouseDown: execute { MAIN_PRG.RobotCommand.trans_x := +1; }
        OnMouseUp: execute { MAIN_PRG.RobotCommand.trans_x := 0; }
    Rectangle (469,445 42x30), "-"
        OnMouseDown: execute { MAIN_PRG.RobotCommand.trans_x := -1; }
        OnMouseUp: execute { MAIN_PRG.RobotCommand.trans_x := 0; }
    Rectangle (417,485 42x30), "+"
        OnMouseDown: execute { MAIN_PRG.RobotCommand.trans_y := +1; }
        OnMouseUp: execute { MAIN_PRG.RobotCommand.trans_y := 0; }
    Rectangle (469,524 42x30), "-"
        OnMouseDown: execute { MAIN_PRG.RobotCommand.trans_z := -1; }
        OnMouseUp: execute { MAIN_PRG.RobotCommand.trans_z := 0; }
    Rectangle (417,524 42x30), "+"
        OnMouseDown: execute { MAIN_PRG.RobotCommand.trans_z := +1; }
        OnMouseUp: execute { MAIN_PRG.RobotCommand.trans_z := 0; }
    Rectangle (417,562 42x30), "+"
        OnMouseDown: execute { MAIN_PRG.RobotCommand.rot_x := +1; }
        OnMouseUp: execute { MAIN_PRG.RobotCommand.rot_x := 0; }
    Rectangle (469,485 42x30), "-"
        OnMouseDown: execute { MAIN_PRG.RobotCommand.trans_y := -1; }
        OnMouseUp: execute { MAIN_PRG.RobotCommand.trans_y := 0; }
    Rectangle (469,562 42x30), "-"
        OnMouseDown: execute { MAIN_PRG.RobotCommand.rot_x := -1; }
        OnMouseUp: execute { MAIN_PRG.RobotCommand.rot_x := 0; }
    Rectangle (417,598 42x30), "+"
        OnMouseDown: execute { MAIN_PRG.RobotCommand.rot_y := +1; }
        OnMouseUp: execute { MAIN_PRG.RobotCommand.rot_y := 0; }
    Rectangle (469,598 42x30), "-"
        OnMouseDown: execute { MAIN_PRG.RobotCommand.rot_y := -1; }
        OnMouseUp: execute { MAIN_PRG.RobotCommand.rot_y := 0; }
    Rectangle (417,638 42x30), "+"
        OnMouseDown: execute { MAIN_PRG.RobotCommand.rot_z := +1; }
        OnMouseUp: execute { MAIN_PRG.RobotCommand.rot_z := 0; }
    Rectangle (469,638 42x30), "-"
        OnMouseDown: execute { MAIN_PRG.RobotCommand.rot_z := -1; }
        OnMouseUp: execute { MAIN_PRG.RobotCommand.rot_z := 0; }
    Slider (281,683 247x47), variable: MAIN_PRG.RobotCommand.tcp_velocity, scale 0..1
    Rectangle (331,404 150x30), "TCP JOG", colour toggle: GVL_OPCUA.RobotCommand.Mode_TCP
        toggle GVL_OPCUA.RobotCommand.Mode_TCP
        OnMouseClick: execute { GVL_OPCUA.RobotCommand.Mode_Axis := FALSE; }
    Rectangle (293,450 104x30), "trans_x"
    Rectangle (293,491 104x30), "trans_y"
    Rectangle (293,526 104x30), "trans_z"
    Rectangle (293,564 104x30), "rot_x"
    Rectangle (293,603 104x30), "rot_y"
    Rectangle (293,638 104x30), "rot_z"
    Rectangle (114,790 210x30), "Info: guter Wert für Velocity: 0.2 - 0.35"
    Rectangle (112,757 509x28), "Wen .n Arm in Singularität feststeckt -> aus Singularität rausfahren mit Joint Jog"
    Rectangle (270,361 97x19), "Status Code"
    Rectangle (375,361 49x19), "%i", text variable: MAIN_PRG.RobotCommand.status
    Rectangle (434,361 94x19), "%s", text variable: MAIN_PRG.Status_Servo
    Rectangle (19,352 95x19), "Translation"
    RoundedRectangle (357,805 264x29), "Skalierungsfaktor für maximale Geschwindigkeit"
END_VISUALIZATION

// Device/Application/VISU_Auto
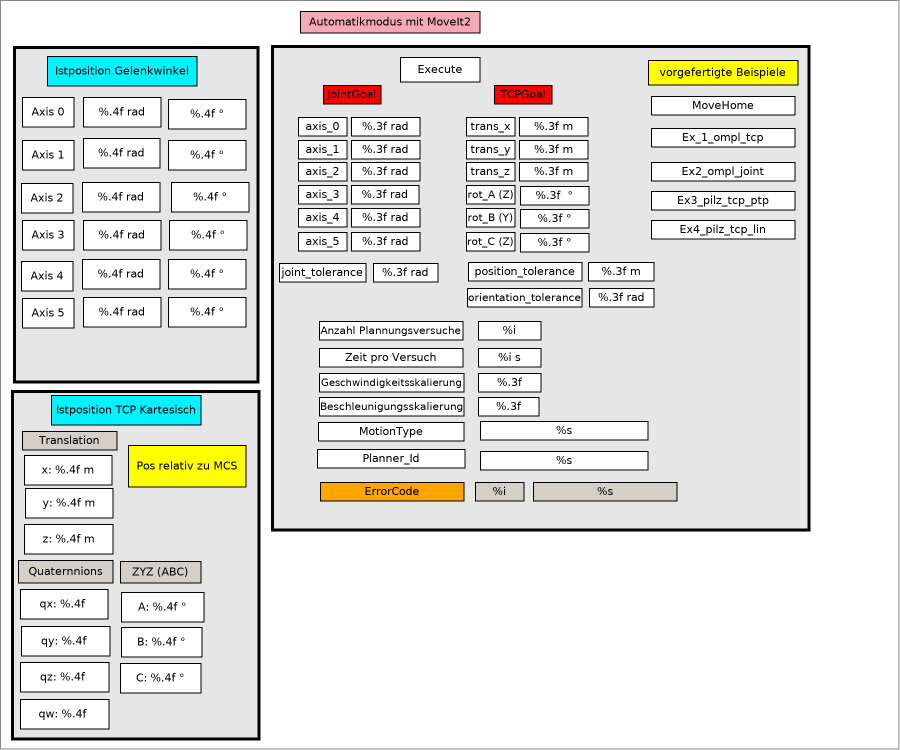
VISUALIZATION VISU_Auto  // 900x750
    Rectangle (271,45 539x486)
    Rectangle (298,117 49x19), "axis_0"
    Rectangle (298,140 49x19), "axis_1"
    Rectangle (298,162 49x19), "axis_2"
    Rectangle (298,185 49x19), "axis_3"
    Rectangle (298,208 49x19), "axis_4"
    Rectangle (298,232 49x19), "axis_5"
    Rectangle (351,117 69x19), "%.3f rad", text variable: MAIN_PRG.RobotAction.axis_0
        OnMouseClick: write the text variable via Default
    Rectangle (351,140 69x19), "%.3f rad", text variable: MAIN_PRG.RobotAction.axis_1
        OnMouseClick: write the text variable via Default
    Rectangle (351,162 69x19), "%.3f rad", text variable: MAIN_PRG.RobotAction.axis_2
        OnMouseClick: write the text variable via Default
    Rectangle (351,185 68x19), "%.3f rad", text variable: MAIN_PRG.RobotAction.axis_3
        OnMouseClick: write the text variable via Default
    Rectangle (351,208 69x19), "%.3f rad", text variable: MAIN_PRG.RobotAction.axis_4
        OnMouseClick: write the text variable via Default
    Rectangle (351,232 69x19), "%.3f rad", text variable: MAIN_PRG.RobotAction.axis_5
        OnMouseClick: write the text variable via Default
    Rectangle (466,117 49x19), "trans_x"
    Rectangle (466,140 49x19), "trans_y"
    Rectangle (466,162 49x19), "trans_z"
    Rectangle (519,117 69x19), "%.3f m", text variable: MAIN_PRG.RobotAction.trans_x
        OnMouseClick: write the text variable via Default
    Rectangle (519,140 69x19), "%.3f m", text variable: MAIN_PRG.RobotAction.trans_y
        OnMouseClick: write the text variable via Default
    Rectangle (519,162 69x19), "%.3f m", text variable: MAIN_PRG.RobotAction.trans_z
        OnMouseClick: write the text variable via Default
    Rectangle (400,57 80x25), "Execute"
        tap GVL_OPCUA.Execute
    Rectangle (323,85 58x19), "JointGoal", colour toggle: MAIN_PRG.RobotAction.Joint_Goal
        toggle MAIN_PRG.RobotAction.Joint_Goal
    Rectangle (494,85 58x19), "TCPGoal", colour toggle: MAIN_PRG.RobotAction.TCP_Goal
        toggle MAIN_PRG.RobotAction.TCP_Goal
    Rectangle (319,321 144x19), "Anzahl Plannungsversuche"
    Rectangle (319,348 144x19), "Zeit pro Versuch"
    Rectangle (319,373 145x19), "Geschwindigkeitsskalierung"
    Rectangle (319,397 145x19), "Beschleunigungsskalierung"
    Rectangle (468,262 114x19), "position_tolerance"
    Rectangle (467,288 115x19), "orientation_tolerance"
    Rectangle (478,321 63x19), "%i", text variable: MAIN_PRG.RobotAction.num_planning_attempts
        OnMouseClick: write the text variable via Default
    Rectangle (478,348 63x19), "%i s", text variable: MAIN_PRG.RobotAction.allowed_planning_time
        OnMouseClick: write the text variable via Default
    Rectangle (478,373 63x19), "%.3f", text variable: MAIN_PRG.RobotAction.max_velocity_scaling
        OnMouseClick: write the text variable via Default
    Rectangle (478,397 61x19), "%.3f", text variable: MAIN_PRG.RobotAction.max_acceleration_scaling
        OnMouseClick: write the text variable via Default
    Rectangle (588,262 66x19), "%.3f m", text variable: MAIN_PRG.RobotAction.position_tolerance
        OnMouseClick: write the text variable via Default
    Rectangle (589,288 65x19), "%.3f rad", text variable: MAIN_PRG.RobotAction.orientation_tolerance
        OnMouseClick: write the text variable via Default
    Rectangle (318,422 146x19), "MotionType"
    Rectangle (317,449 148x19), "Planner_Id"
    Rectangle (320,482 144x19), "ErrorCode"
    Rectangle (475,482 49x19), "%i", text variable: MAIN_PRG.RobotAction.error_code
    Rectangle (480,421 168x19), "%s", text variable: MAIN_PRG.RobotAction.Motion_Type
        OnMouseClick: write the text variable via Default
    Rectangle (480,451 168x19), "%s", text variable: MAIN_PRG.RobotAction.Planner_ID
        OnMouseClick: write the text variable via Default
    Rectangle (651,96 144x19), "MoveHome"
        tap MAIN_PRG.xMoveHome
    Rectangle (533,482 144x19), "%s", text variable: MAIN_PRG.Status_Error_Codes_Action
    Rectangle (651,128 144x19), "Ex_1_ompl_tcp"
        tap MAIN_PRG.xEx1_ompl_tcp
    Rectangle (651,162 144x19), "Ex2_ompl_joint"
        tap MAIN_PRG.xEx2_ompl_joint
    Rectangle (651,191 144x19), "Ex3_pilz_tcp_ptp"
        tap MAIN_PRG.xEx3_pilz_tcp_ptp
    Rectangle (651,220 144x19), "Ex4_pilz_tcp_lin"
        tap MAIN_PRG.xEx4_pilz_tcp_lin
    RoundedRectangle (648,60 150x25), "vorgefertigte Beispiele"
    Rectangle (466,185 49x19), "rot_A (Z)"
    Rectangle (466,208 49x19), "rot_B (Y)"
    Rectangle (466,232 49x19), "rot_C (Z)"
    Rectangle (520,186 69x19), "%.3f °", text variable: GVL_OPCUA.rot_A
        OnMouseClick: write the text variable via Default
    Rectangle (520,209 69x19), "%.3f °", text variable: GVL_OPCUA.rot_B
        OnMouseClick: write the text variable via Default
    Rectangle (520,233 69x19), "%.3f °", text variable: GVL_OPCUA.rot_C
        OnMouseClick: write the text variable via Default
    Rectangle (279,263 87x19), "joint_tolerance"
    Rectangle (373,263 65x19), "%.3f rad", text variable: MAIN_PRG.RobotAction.joint_tolerance
        OnMouseClick: write the text variable via Default
    Rectangle (11,390 249x350)
    Rectangle (13,46 246x337)
    Rectangle (47,56 150x30), "Istposition Gelenkwinkel"
    Rectangle (51,395 150x30), "Istposition TCP Kartesisch"
    Rectangle (24,455 88x30), "x: %.4f m", text variable: MAIN_PRG.RobotStatus.tcp_pose.trans_x
    Rectangle (25,488 88x30), "y: %.4f m", text variable: MAIN_PRG.RobotStatus.tcp_pose.trans_y
    Rectangle (24,524 89x30), "z: %.4f m", text variable: MAIN_PRG.RobotStatus.tcp_pose.trans_z
    Rectangle (20,589 88x30), "qx: %.4f", text variable: MAIN_PRG.RobotStatus.tcp_pose.rot_x
    Rectangle (21,626 89x30), "qy: %.4f", text variable: MAIN_PRG.RobotStatus.tcp_pose.rot_y
    Rectangle (20,662 89x30), "qz: %.4f", text variable: MAIN_PRG.RobotStatus.tcp_pose.rot_z
    Rectangle (20,699 89x30), "qw: %.4f", text variable: MAIN_PRG.RobotStatus.tcp_pose.rot_w
    Rectangle (83,97 78x30), "%.4f rad", text variable: MAIN_PRG.RobotStatus.axis_pose.axis_0
    Rectangle (83,138 77x30), "%.4f rad", text variable: MAIN_PRG.RobotStatus.axis_pose.axis_1
    Rectangle (82,182 78x30), "%.4f rad", text variable: MAIN_PRG.RobotStatus.axis_pose.axis_2
    Rectangle (83,220 78x30), "%.4f rad", text variable: MAIN_PRG.RobotStatus.axis_pose.axis_3
    Rectangle (82,259 78x30), "%.4f rad", text variable: MAIN_PRG.RobotStatus.axis_pose.axis_4
    Rectangle (83,297 78x30), "%.4f rad", text variable: MAIN_PRG.RobotStatus.axis_pose.axis_5
    Rectangle (168,99 78x30), "%.4f °", text variable: MAIN_PRG.RobotStatus.axis_pose.axis_0 *(180.0/GVL_OPCUA.PI)
    Rectangle (168,140 78x30), "%.4f °", text variable: MAIN_PRG.RobotStatus.axis_pose.axis_1 *(180.0/GVL_OPCUA.PI)
    Rectangle (171,182 78x30), "%.4f °", text variable: MAIN_PRG.RobotStatus.axis_pose.axis_2 *(180.0/GVL_OPCUA.PI)
    Rectangle (169,220 78x30), "%.4f °", text variable: MAIN_PRG.RobotStatus.axis_pose.axis_3 *(180.0/GVL_OPCUA.PI)
    Rectangle (168,259 78x30), "%.4f °", text variable: MAIN_PRG.RobotStatus.axis_pose.axis_4 *(180.0/GVL_OPCUA.PI)
    Rectangle (168,297 78x30), "%.4f °", text variable: MAIN_PRG.RobotStatus.axis_pose.axis_5 *(180.0/GVL_OPCUA.PI)
    Rectangle (121,592 83x30), "A: %.4f °", text variable: MAIN_PRG.Status_Quat_to_ZYZ.euler.A
    Rectangle (121,627 81x30), "B: %.4f °", text variable: MAIN_PRG.Status_Quat_to_ZYZ.euler.B
    Rectangle (120,663 81x30), "C: %.4f °", text variable: MAIN_PRG.Status_Quat_to_ZYZ.euler.C
    Rectangle (120,561 81x22), "ZYZ (ABC)"
    Rectangle (18,560 95x23), "Quaternnions"
    Rectangle (22,97 52x30), "Axis 0"
    Rectangle (22,140 52x30), "Axis 1"
    Rectangle (21,183 52x30), "Axis 2"
    Rectangle (22,220 52x30), "Axis 3"
    Rectangle (21,261 52x30), "Axis 4"
    Rectangle (22,298 52x30), "Axis 5"
    RoundedRectangle (128,445 118x42), "Pos relativ zu MCS"
    Rectangle (22,431 95x19), "Translation"
    Rectangle (300,11 180x22), "Automatikmodus mit MoveIt2"
END_VISUALIZATION

// Device/Application/VISU_Startseite
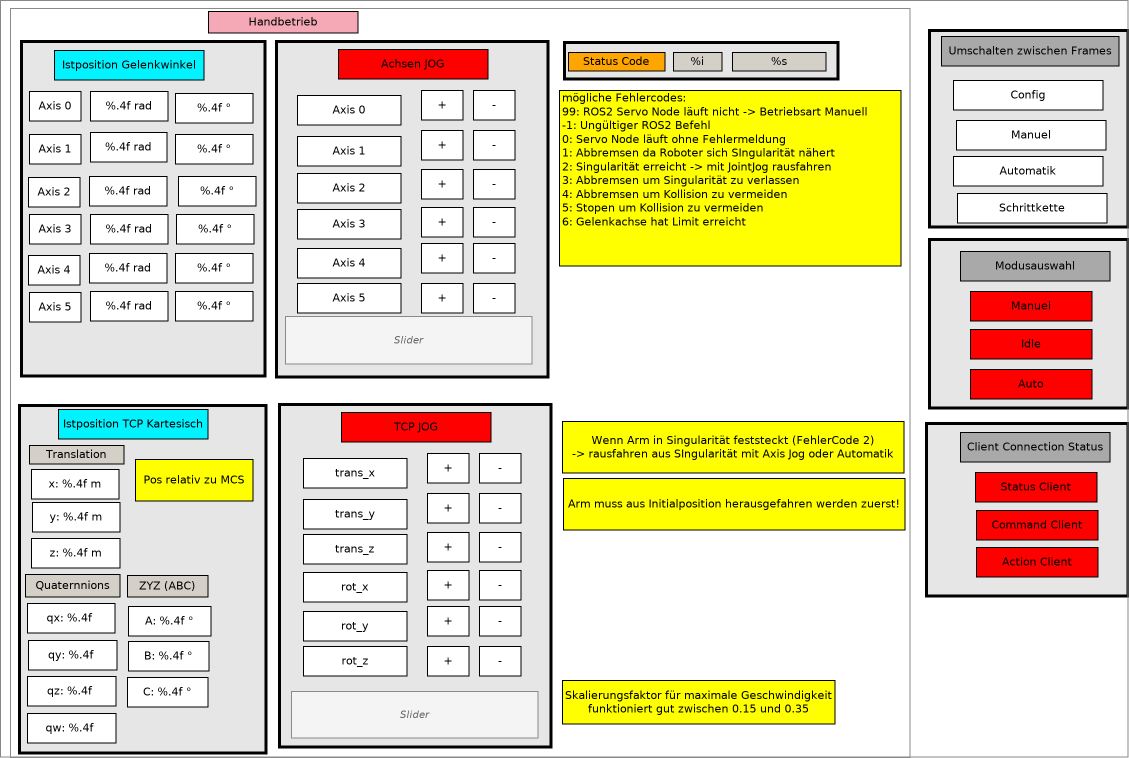
VISUALIZATION VISU_Startseite  // 1129x758
    Rectangle (928,29 201x199)
    Frame (10,8 900x750)
        shows VISU_Manuell()
        shows VISU_Konfig()
        shows VISU_Auto()
        shows VISU_Schrittkette()
    Rectangle (953,80 150x30), "Config"
        OnMouseClick: FrameSelectionChange Selection=SelectedFrame=848abb15-4fea-4ce4-a60a-73a186e6a183, Selection=1, GlobSel=AssignType=Directly, SelType=Locally, SelectionStep=SelectedAction=SwitchNext
    Rectangle (956,120 150x30), "Manuel"
        OnMouseClick: FrameSelectionChange Selection=SelectedFrame=848abb15-4fea-4ce4-a60a-73a186e6a183, GlobSel=AssignType=Directly, SelType=Locally, SelectionStep=SelectedAction=SwitchNext
    Rectangle (953,156 150x30), "Automatik"
        OnMouseClick: FrameSelectionChange Selection=SelectedFrame=848abb15-4fea-4ce4-a60a-73a186e6a183, Selection=2, GlobSel=AssignType=Directly, SelType=Locally, SelectionStep=SelectedAction=SwitchNext
    Rectangle (941,36 178x30), "Umschalten zwischen Frames"
    Rectangle (928,238 201x171)
    Rectangle (960,251 150x30), "Modusauswahl"
    Rectangle (970,291 122x30), "Manuel", colour toggle: MAIN_PRG.Modes.MANUEL
        toggle MAIN_PRG.Modes.SEL_MAN p2164770859=TRUE
    Rectangle (970,369 122x30), "Auto", colour toggle: MAIN_PRG.Modes.AUTO
        toggle MAIN_PRG.Modes.SEL_AUTO p2164770859=TRUE
    Rectangle (970,329 122x30), "Idle", colour toggle: MAIN_PRG.Modes.IDLE
    Rectangle (925,422 204x175)
    Rectangle (960,432 150x30), "Client Connection Status"
    Rectangle (975,472 122x30), "Status Client", colour toggle: MAIN_PRG.RobotStatus.client_connected
    Rectangle (976,547 122x30), "Action Client", colour toggle: MAIN_PRG.RobotAction.client_connected
    Rectangle (976,510 122x30), "Command Client", colour toggle: MAIN_PRG.RobotCommand.client_connected
    Rectangle (957,193 150x30), "Schrittkette"
        OnMouseClick: FrameSelectionChange Selection=SelectedFrame=848abb15-4fea-4ce4-a60a-73a186e6a183, Selection=3, GlobSel=AssignType=Directly, SelType=Locally, SelectionStep=SelectedAction=SwitchNext
END_VISUALIZATION

// Device/Application/VISU_Manuell
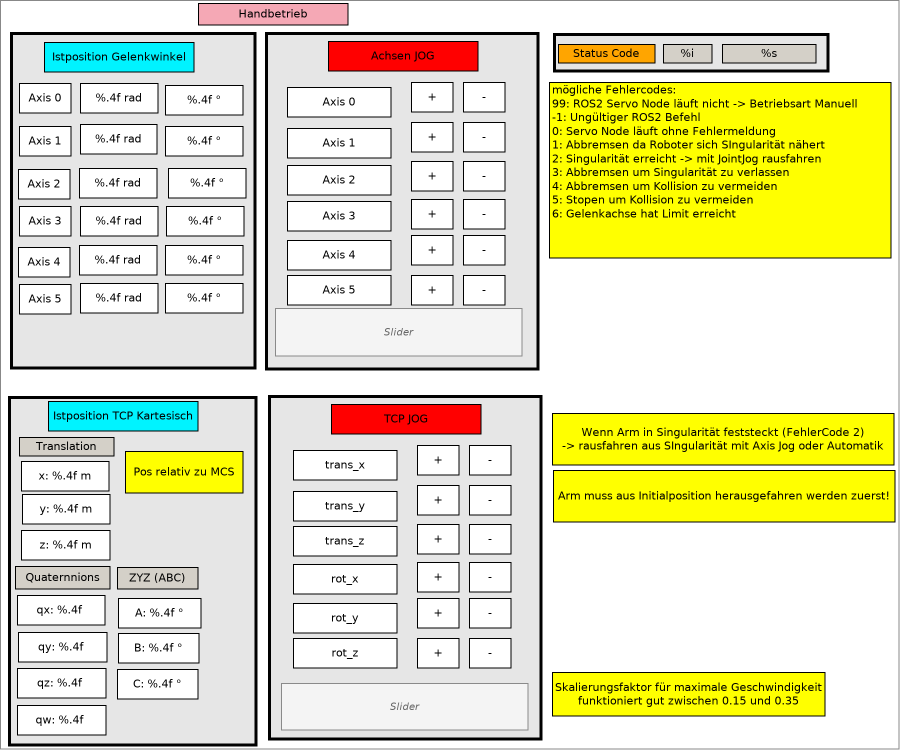
VISUALIZATION VISU_Manuell  // 900x750
    Rectangle (553,33 276x39)
    Rectangle (265,32 274x338)
    Rectangle (8,396 249x350)
    Rectangle (10,32 246x337)
    Rectangle (44,42 150x30), "Istposition Gelenkwinkel"
    Rectangle (48,401 150x30), "Istposition TCP Kartesisch"
    Rectangle (21,461 88x30), "x: %.4f m", text variable: MAIN_PRG.RobotStatus.tcp_pose.trans_x
    Rectangle (22,494 88x30), "y: %.4f m", text variable: MAIN_PRG.RobotStatus.tcp_pose.trans_y
    Rectangle (21,530 89x30), "z: %.4f m", text variable: MAIN_PRG.RobotStatus.tcp_pose.trans_z
    Rectangle (17,595 88x30), "qx: %.4f", text variable: MAIN_PRG.RobotStatus.tcp_pose.rot_x
    Rectangle (18,632 89x30), "qy: %.4f", text variable: MAIN_PRG.RobotStatus.tcp_pose.rot_y
    Rectangle (17,668 89x30), "qz: %.4f", text variable: MAIN_PRG.RobotStatus.tcp_pose.rot_z
    Rectangle (17,705 89x30), "qw: %.4f", text variable: MAIN_PRG.RobotStatus.tcp_pose.rot_w
    Rectangle (411,82 42x30), "+"
        OnMouseDown: execute { MAIN_PRG.RobotCommand.axis_0 := +1; }
        OnMouseUp: execute { MAIN_PRG.RobotCommand.axis_0 := 0; }
    Rectangle (463,82 42x30), "-"
        OnMouseDown: execute { MAIN_PRG.RobotCommand.axis_0 := -1; }
        OnMouseUp: execute { MAIN_PRG.RobotCommand.axis_0 := 0; }
    Rectangle (411,122 42x30), "+"
        OnMouseDown: execute { MAIN_PRG.RobotCommand.axis_1 := +1; }
        OnMouseUp: execute { MAIN_PRG.RobotCommand.axis_1 := 0; }
    Rectangle (463,161 42x30), "-"
        OnMouseDown: execute { MAIN_PRG.RobotCommand.axis_2 := -1; }
        OnMouseUp: execute { MAIN_PRG.RobotCommand.axis_2 := 0; }
    Rectangle (411,161 42x30), "+"
        OnMouseDown: execute { MAIN_PRG.RobotCommand.axis_2 := +1; }
        OnMouseUp: execute { MAIN_PRG.RobotCommand.axis_2 := 0; }
    Rectangle (411,199 42x30), "+"
        OnMouseDown: execute { MAIN_PRG.RobotCommand.axis_3 := +1; }
        OnMouseUp: execute { MAIN_PRG.RobotCommand.axis_3 := 0; }
    Rectangle (463,122 42x30), "-"
        OnMouseDown: execute { MAIN_PRG.RobotCommand.axis_1 := -1; }
        OnMouseUp: execute { MAIN_PRG.RobotCommand.axis_1 := 0; }
    Rectangle (463,199 42x30), "-"
        OnMouseDown: execute { MAIN_PRG.RobotCommand.axis_3 := -1; }
        OnMouseUp: execute { MAIN_PRG.RobotCommand.axis_3 := 0; }
    Rectangle (411,235 42x30), "+"
        OnMouseDown: execute { MAIN_PRG.RobotCommand.axis_4 := +1; }
        OnMouseUp: execute { MAIN_PRG.RobotCommand.axis_4 := 0; }
    Rectangle (463,235 42x30), "-"
        OnMouseDown: execute { MAIN_PRG.RobotCommand.axis_4 := -1; }
        OnMouseUp: execute { MAIN_PRG.RobotCommand.axis_4 := 0; }
    Rectangle (411,275 42x30), "+"
        OnMouseDown: execute { MAIN_PRG.RobotCommand.axis_5 := +1; }
        OnMouseUp: execute { MAIN_PRG.RobotCommand.axis_5 := 0; }
    Rectangle (463,275 42x30), "-"
        OnMouseDown: execute { MAIN_PRG.RobotCommand.axis_5 := -1; }
        OnMouseUp: execute { MAIN_PRG.RobotCommand.axis_5 := 0; }
    Slider (275,308 247x48), variable: MAIN_PRG.RobotCommand.axis_velocity, scale 0..1
    Rectangle (80,83 78x30), "%.4f rad", text variable: MAIN_PRG.RobotStatus.axis_pose.axis_0
    Rectangle (80,124 77x30), "%.4f rad", text variable: MAIN_PRG.RobotStatus.axis_pose.axis_1
    Rectangle (79,168 78x30), "%.4f rad", text variable: MAIN_PRG.RobotStatus.axis_pose.axis_2
    Rectangle (80,206 78x30), "%.4f rad", text variable: MAIN_PRG.RobotStatus.axis_pose.axis_3
    Rectangle (79,245 78x30), "%.4f rad", text variable: MAIN_PRG.RobotStatus.axis_pose.axis_4
    Rectangle (80,283 78x30), "%.4f rad", text variable: MAIN_PRG.RobotStatus.axis_pose.axis_5
    Rectangle (328,41 150x30), "Achsen JOG", colour toggle: GVL_OPCUA.RobotCommand.Mode_Axis
        toggle GVL_OPCUA.RobotCommand.Mode_Axis
        OnMouseClick: execute { GVL_OPCUA.RobotCommand.Mode_TCP := FALSE; }
    Rectangle (165,85 78x30), "%.4f °", text variable: MAIN_PRG.RobotStatus.axis_pose.axis_0 *(180.0/GVL_OPCUA.PI)
    Rectangle (165,126 78x30), "%.4f °", text variable: MAIN_PRG.RobotStatus.axis_pose.axis_1 *(180.0/GVL_OPCUA.PI)
    Rectangle (168,168 78x30), "%.4f °", text variable: MAIN_PRG.RobotStatus.axis_pose.axis_2 *(180.0/GVL_OPCUA.PI)
    Rectangle (166,206 78x30), "%.4f °", text variable: MAIN_PRG.RobotStatus.axis_pose.axis_3 *(180.0/GVL_OPCUA.PI)
    Rectangle (165,245 78x30), "%.4f °", text variable: MAIN_PRG.RobotStatus.axis_pose.axis_4 *(180.0/GVL_OPCUA.PI)
    Rectangle (165,283 78x30), "%.4f °", text variable: MAIN_PRG.RobotStatus.axis_pose.axis_5 *(180.0/GVL_OPCUA.PI)
    Rectangle (118,598 83x30), "A: %.4f °", text variable: MAIN_PRG.Status_Quat_to_ZYZ.euler.A
    Rectangle (118,633 81x30), "B: %.4f °", text variable: MAIN_PRG.Status_Quat_to_ZYZ.euler.B
    Rectangle (117,669 81x30), "C: %.4f °", text variable: MAIN_PRG.Status_Quat_to_ZYZ.euler.C
    Rectangle (117,567 81x22), "ZYZ (ABC)"
    Rectangle (15,566 95x23), "Quaternnions"
    Rectangle (287,87 104x30), "Axis 0"
    Rectangle (287,128 104x30), "Axis 1"
    Rectangle (287,165 104x30), "Axis 2"
    Rectangle (287,201 104x30), "Axis 3"
    Rectangle (287,240 104x30), "Axis 4"
    Rectangle (287,275 104x30), "Axis 5"
    Rectangle (19,83 52x30), "Axis 0"
    Rectangle (19,126 52x30), "Axis 1"
    Rectangle (18,169 52x30), "Axis 2"
    Rectangle (19,206 52x30), "Axis 3"
    Rectangle (18,247 52x30), "Axis 4"
    Rectangle (19,284 52x30), "Axis 5"
    RoundedRectangle (125,451 118x42), "Pos relativ zu MCS"
    Rectangle (268,395 274x345)
    Rectangle (417,445 42x30), "+"
        OnMouseDown: execute { MAIN_PRG.RobotCommand.trans_x := +1; }
        OnMouseUp: execute { MAIN_PRG.RobotCommand.trans_x := 0; }
    Rectangle (469,445 42x30), "-"
        OnMouseDown: execute { MAIN_PRG.RobotCommand.trans_x := -1; }
        OnMouseUp: execute { MAIN_PRG.RobotCommand.trans_x := 0; }
    Rectangle (417,485 42x30), "+"
        OnMouseDown: execute { MAIN_PRG.RobotCommand.trans_y := +1; }
        OnMouseUp: execute { MAIN_PRG.RobotCommand.trans_y := 0; }
    Rectangle (469,524 42x30), "-"
        OnMouseDown: execute { MAIN_PRG.RobotCommand.trans_z := -1; }
        OnMouseUp: execute { MAIN_PRG.RobotCommand.trans_z := 0; }
    Rectangle (417,524 42x30), "+"
        OnMouseDown: execute { MAIN_PRG.RobotCommand.trans_z := +1; }
        OnMouseUp: execute { MAIN_PRG.RobotCommand.trans_z := 0; }
    Rectangle (417,562 42x30), "+"
        OnMouseDown: execute { MAIN_PRG.RobotCommand.rot_x := +1; }
        OnMouseUp: execute { MAIN_PRG.RobotCommand.rot_x := 0; }
    Rectangle (469,485 42x30), "-"
        OnMouseDown: execute { MAIN_PRG.RobotCommand.trans_y := -1; }
        OnMouseUp: execute { MAIN_PRG.RobotCommand.trans_y := 0; }
    Rectangle (469,562 42x30), "-"
        OnMouseDown: execute { MAIN_PRG.RobotCommand.rot_x := -1; }
        OnMouseUp: execute { MAIN_PRG.RobotCommand.rot_x := 0; }
    Rectangle (417,598 42x30), "+"
        OnMouseDown: execute { MAIN_PRG.RobotCommand.rot_y := +1; }
        OnMouseUp: execute { MAIN_PRG.RobotCommand.rot_y := 0; }
    Rectangle (469,598 42x30), "-"
        OnMouseDown: execute { MAIN_PRG.RobotCommand.rot_y := -1; }
        OnMouseUp: execute { MAIN_PRG.RobotCommand.rot_y := 0; }
    Rectangle (417,638 42x30), "+"
        OnMouseDown: execute { MAIN_PRG.RobotCommand.rot_z := +1; }
        OnMouseUp: execute { MAIN_PRG.RobotCommand.rot_z := 0; }
    Rectangle (469,638 42x30), "-"
        OnMouseDown: execute { MAIN_PRG.RobotCommand.rot_z := -1; }
        OnMouseUp: execute { MAIN_PRG.RobotCommand.rot_z := 0; }
    Slider (281,683 247x47), variable: MAIN_PRG.RobotCommand.tcp_velocity, scale 0..1
    Rectangle (331,404 150x30), "TCP JOG", colour toggle: GVL_OPCUA.RobotCommand.Mode_TCP
        toggle GVL_OPCUA.RobotCommand.Mode_TCP
        OnMouseClick: execute { GVL_OPCUA.RobotCommand.Mode_Axis := FALSE; }
    Rectangle (293,450 104x30), "trans_x"
    Rectangle (293,491 104x30), "trans_y"
    Rectangle (293,526 104x30), "trans_z"
    Rectangle (293,564 104x30), "rot_x"
    Rectangle (293,603 104x30), "rot_y"
    Rectangle (293,638 104x30), "rot_z"
    Rectangle (558,44 97x19), "Status Code"
    Rectangle (663,44 49x19), "%i", text variable: MAIN_PRG.RobotCommand.status
    Rectangle (722,44 94x19), "%s", text variable: MAIN_PRG.Status_Servo
    Rectangle (19,437 95x19), "Translation"
    RoundedRectangle (552,672 273x44), "Skalierungsfaktor für maximale Geschwindigkeit funktioniert gut zwischen 0.15 und 0.35"
    Rectangle (198,3 150x22), "Handbetrieb"
    RoundedRectangle (552,413 342x52), "Wenn Arm in Singularität feststeckt (FehlerCode 2) -> rausfahren aus SIngularität mit Axis Jog oder Automatik"
    RoundedRectangle (549,82 342x176), "mögliche Fehlercodes: 99: ROS2 Servo Node läuft nicht -> Betriebsart Manuell -1: Ungültiger ROS2 Befehl 0: Servo Node läuft ohne Fehlermeldung 1: Abbremsen da Roboter sich SIngularität nähert 2: Singularität erreicht -> mit JointJog rausfahren 3: Abbremsen um Singularität zu verlassen 4: Abbremsen um Kollision zu vermeiden 5: Stopen um Kollision zu vermeiden 6: Gelenkachse hat Limit erreicht"
    RoundedRectangle (553,470 342x52), "Arm muss aus Initialposition herausgefahren werden zuerst!"
END_VISUALIZATION

// Device/Application/VISU_Konfig
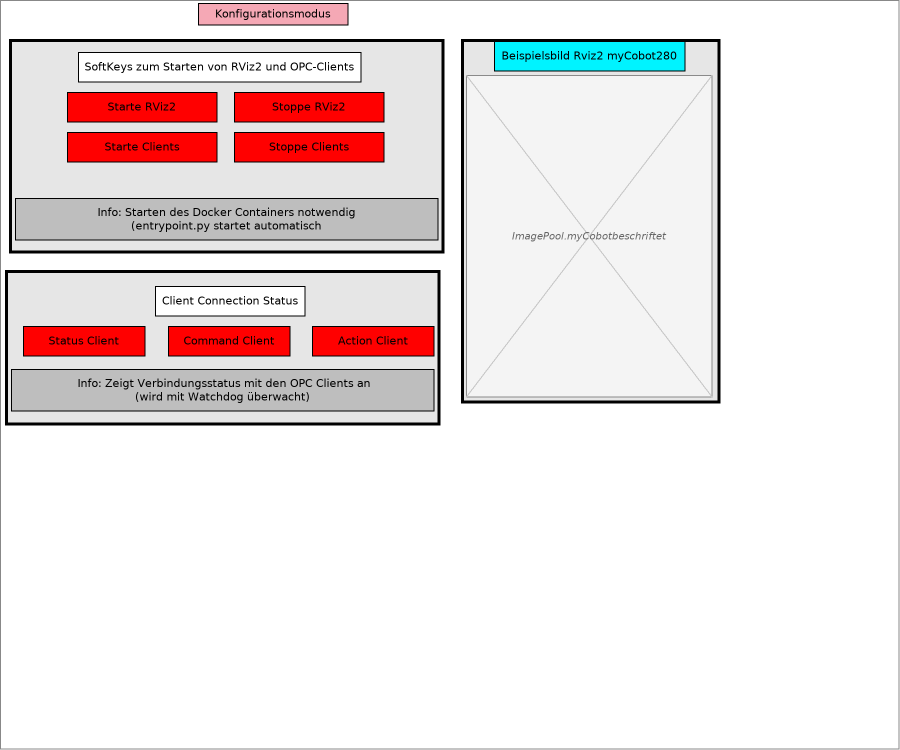
VISUALIZATION VISU_Konfig  // 900x750
    Rectangle (198,3 150x22), "Konfigurationsmodus"
    Rectangle (461,39 259x364)
    Rectangle (9,39 435x214)
    Rectangle (67,92 150x30), "Starte RViz2"
        toggle GVL_OPCUA.Start_RViz2
    Rectangle (67,132 150x30), "Starte Clients"
        toggle GVL_OPCUA.Start_OPCClients
    Rectangle (234,132 150x30), "Stoppe Clients"
        toggle GVL_OPCUA.Stop_OPC_Clients
    Rectangle (234,92 150x30), "Stoppe RViz2"
        toggle GVL_OPCUA.Stop_RViz2
    Image (466,75 246x322), image: ImagePool.myCobotbeschriftet
    Rectangle (494,41 191x30), "Beispielsbild Rviz2 myCobot280"
    Rectangle (78,52 283x30), "SoftKeys zum Starten von RViz2 und OPC-Clients"
    Rectangle (15,198 423x42), "Info: Starten des Docker Containers notwendig (entrypoint.py startet automatisch"
    Rectangle (5,270 435x155)
    Rectangle (155,286 150x30), "Client Connection Status"
    Rectangle (23,326 122x30), "Status Client", colour toggle: MAIN_PRG.RobotStatus.client_connected
    Rectangle (312,326 122x30), "Action Client", colour toggle: MAIN_PRG.RobotAction.client_connected
    Rectangle (168,326 122x30), "Command Client", colour toggle: MAIN_PRG.RobotCommand.client_connected
    Rectangle (11,369 423x42), "Info: Zeigt Verbindungsstatus mit den OPC Clients an (wird mit Watchdog überwacht)"
END_VISUALIZATION

// Device/Application/VISU_Schrittkette
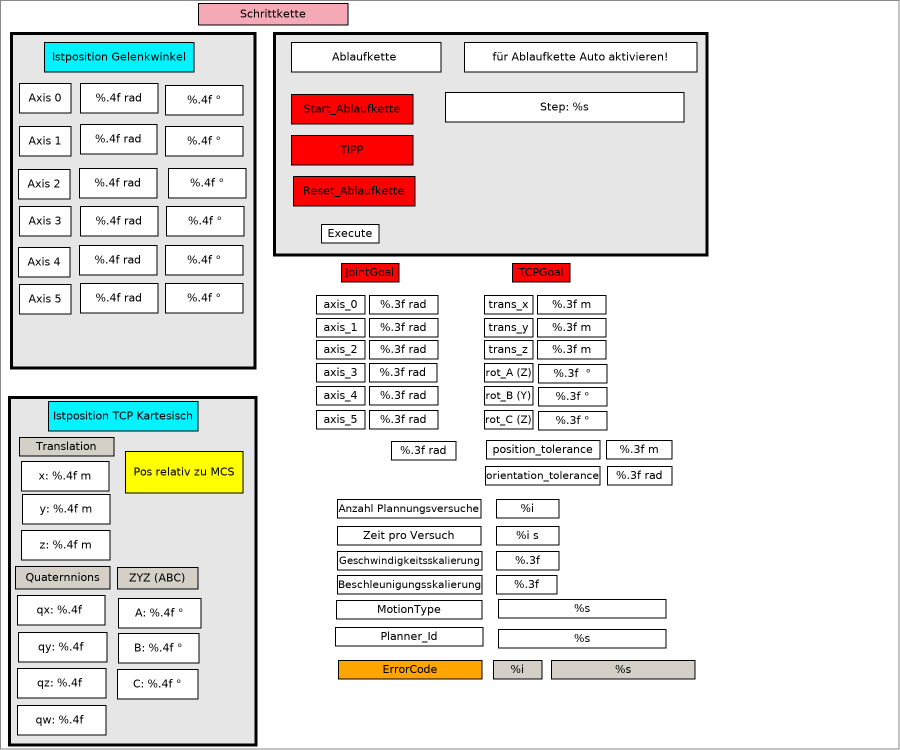
VISUALIZATION VISU_Schrittkette  // 900x750
    Rectangle (273,32 435x224)
    Rectangle (291,42 150x30), "Ablaufkette"
    Rectangle (291,135 122x30), "TIPP", colour toggle: MAIN_PRG.RobotStatus.client_connected
        tap GVL_OPCUA.TIPP
    Rectangle (291,94 122x30), "Start_Ablaufkette", colour toggle: MAIN_PRG.RobotStatus.client_connected
        tap GVL_OPCUA.Start_Ablaufkette
    Rectangle (445,92 239x30), "Step: %s", text variable: Ablaufkette.SFCCurrentStep
    Rectangle (464,42 233x30), "für Ablaufkette Auto aktivieren!"
    Rectangle (293,176 122x30), "Reset_Ablaufkette", colour toggle: MAIN_PRG.RobotStatus.client_connected
        tap GVL_OPCUA.Reset_Ablaufkette
    Rectangle (321,224 58x19), "Execute"
        tap GVL_OPCUA.Execute
    Rectangle (8,396 249x350)
    Rectangle (10,32 246x337)
    Rectangle (44,42 150x30), "Istposition Gelenkwinkel"
    Rectangle (48,401 150x30), "Istposition TCP Kartesisch"
    Rectangle (21,461 88x30), "x: %.4f m", text variable: MAIN_PRG.RobotStatus.tcp_pose.trans_x
    Rectangle (22,494 88x30), "y: %.4f m", text variable: MAIN_PRG.RobotStatus.tcp_pose.trans_y
    Rectangle (21,530 89x30), "z: %.4f m", text variable: MAIN_PRG.RobotStatus.tcp_pose.trans_z
    Rectangle (17,595 88x30), "qx: %.4f", text variable: MAIN_PRG.RobotStatus.tcp_pose.rot_x
    Rectangle (18,632 89x30), "qy: %.4f", text variable: MAIN_PRG.RobotStatus.tcp_pose.rot_y
    Rectangle (17,668 89x30), "qz: %.4f", text variable: MAIN_PRG.RobotStatus.tcp_pose.rot_z
    Rectangle (17,705 89x30), "qw: %.4f", text variable: MAIN_PRG.RobotStatus.tcp_pose.rot_w
    Rectangle (80,83 78x30), "%.4f rad", text variable: MAIN_PRG.RobotStatus.axis_pose.axis_0
    Rectangle (80,124 77x30), "%.4f rad", text variable: MAIN_PRG.RobotStatus.axis_pose.axis_1
    Rectangle (79,168 78x30), "%.4f rad", text variable: MAIN_PRG.RobotStatus.axis_pose.axis_2
    Rectangle (80,206 78x30), "%.4f rad", text variable: MAIN_PRG.RobotStatus.axis_pose.axis_3
    Rectangle (79,245 78x30), "%.4f rad", text variable: MAIN_PRG.RobotStatus.axis_pose.axis_4
    Rectangle (80,283 78x30), "%.4f rad", text variable: MAIN_PRG.RobotStatus.axis_pose.axis_5
    Rectangle (165,85 78x30), "%.4f °", text variable: MAIN_PRG.RobotStatus.axis_pose.axis_0 *(180.0/GVL_OPCUA.PI)
    Rectangle (165,126 78x30), "%.4f °", text variable: MAIN_PRG.RobotStatus.axis_pose.axis_1 *(180.0/GVL_OPCUA.PI)
    Rectangle (168,168 78x30), "%.4f °", text variable: MAIN_PRG.RobotStatus.axis_pose.axis_2 *(180.0/GVL_OPCUA.PI)
    Rectangle (166,206 78x30), "%.4f °", text variable: MAIN_PRG.RobotStatus.axis_pose.axis_3 *(180.0/GVL_OPCUA.PI)
    Rectangle (165,245 78x30), "%.4f °", text variable: MAIN_PRG.RobotStatus.axis_pose.axis_4 *(180.0/GVL_OPCUA.PI)
    Rectangle (165,283 78x30), "%.4f °", text variable: MAIN_PRG.RobotStatus.axis_pose.axis_5 *(180.0/GVL_OPCUA.PI)
    Rectangle (118,598 83x30), "A: %.4f °", text variable: MAIN_PRG.Status_Quat_to_ZYZ.euler.A
    Rectangle (118,633 81x30), "B: %.4f °", text variable: MAIN_PRG.Status_Quat_to_ZYZ.euler.B
    Rectangle (117,669 81x30), "C: %.4f °", text variable: MAIN_PRG.Status_Quat_to_ZYZ.euler.C
    Rectangle (117,567 81x22), "ZYZ (ABC)"
    Rectangle (15,566 95x23), "Quaternnions"
    Rectangle (19,83 52x30), "Axis 0"
    Rectangle (19,126 52x30), "Axis 1"
    Rectangle (18,169 52x30), "Axis 2"
    Rectangle (19,206 52x30), "Axis 3"
    Rectangle (18,247 52x30), "Axis 4"
    Rectangle (19,284 52x30), "Axis 5"
    RoundedRectangle (125,451 118x42), "Pos relativ zu MCS"
    Rectangle (19,437 95x19), "Translation"
    Rectangle (198,3 150x22), "Schrittkette"
    Rectangle (316,295 49x19), "axis_0"
    Rectangle (316,318 49x19), "axis_1"
    Rectangle (316,340 49x19), "axis_2"
    Rectangle (316,363 49x19), "axis_3"
    Rectangle (316,386 49x19), "axis_4"
    Rectangle (316,410 49x19), "axis_5"
    Rectangle (369,295 69x19), "%.3f rad", text variable: MAIN_PRG.RobotAction.axis_0
        OnMouseClick: write the text variable via Default
    Rectangle (369,318 69x19), "%.3f rad", text variable: MAIN_PRG.RobotAction.axis_1
        OnMouseClick: write the text variable via Default
    Rectangle (369,340 69x19), "%.3f rad", text variable: MAIN_PRG.RobotAction.axis_2
        OnMouseClick: write the text variable via Default
    Rectangle (369,363 68x19), "%.3f rad", text variable: MAIN_PRG.RobotAction.axis_3
        OnMouseClick: write the text variable via Default
    Rectangle (369,386 69x19), "%.3f rad", text variable: MAIN_PRG.RobotAction.axis_4
        OnMouseClick: write the text variable via Default
    Rectangle (369,410 69x19), "%.3f rad", text variable: MAIN_PRG.RobotAction.axis_5
        OnMouseClick: write the text variable via Default
    Rectangle (484,295 49x19), "trans_x"
    Rectangle (484,318 49x19), "trans_y"
    Rectangle (484,340 49x19), "trans_z"
    Rectangle (537,295 69x19), "%.3f m", text variable: MAIN_PRG.RobotAction.trans_x
        OnMouseClick: write the text variable via Default
    Rectangle (537,318 69x19), "%.3f m", text variable: MAIN_PRG.RobotAction.trans_y
        OnMouseClick: write the text variable via Default
    Rectangle (537,340 69x19), "%.3f m", text variable: MAIN_PRG.RobotAction.trans_z
        OnMouseClick: write the text variable via Default
    Rectangle (341,263 58x19), "JointGoal", colour toggle: MAIN_PRG.RobotAction.Joint_Goal
        toggle MAIN_PRG.RobotAction.Joint_Goal
    Rectangle (512,263 58x19), "TCPGoal", colour toggle: MAIN_PRG.RobotAction.TCP_Goal
        toggle MAIN_PRG.RobotAction.TCP_Goal
    Rectangle (337,499 144x19), "Anzahl Plannungsversuche"
    Rectangle (337,526 144x19), "Zeit pro Versuch"
    Rectangle (337,551 145x19), "Geschwindigkeitsskalierung"
    Rectangle (337,575 145x19), "Beschleunigungsskalierung"
    Rectangle (486,440 114x19), "position_tolerance"
    Rectangle (485,466 115x19), "orientation_tolerance"
    Rectangle (496,499 63x19), "%i", text variable: MAIN_PRG.RobotAction.num_planning_attempts
        OnMouseClick: write the text variable via Default
    Rectangle (496,526 63x19), "%i s", text variable: MAIN_PRG.RobotAction.allowed_planning_time
        OnMouseClick: write the text variable via Default
    Rectangle (496,551 63x19), "%.3f", text variable: MAIN_PRG.RobotAction.max_velocity_scaling
        OnMouseClick: write the text variable via Default
    Rectangle (496,575 61x19), "%.3f", text variable: MAIN_PRG.RobotAction.max_acceleration_scaling
        OnMouseClick: write the text variable via Default
    Rectangle (606,440 66x19), "%.3f m", text variable: MAIN_PRG.RobotAction.position_tolerance
        OnMouseClick: write the text variable via Default
    Rectangle (607,466 65x19), "%.3f rad", text variable: MAIN_PRG.RobotAction.orientation_tolerance
        OnMouseClick: write the text variable via Default
    Rectangle (336,600 146x19), "MotionType"
    Rectangle (335,627 148x19), "Planner_Id"
    Rectangle (338,660 144x19), "ErrorCode"
    Rectangle (493,660 49x19), "%i", text variable: MAIN_PRG.RobotAction.error_code
    Rectangle (498,599 168x19), "%s", text variable: MAIN_PRG.RobotAction.Motion_Type
        OnMouseClick: write the text variable via Default
    Rectangle (498,629 168x19), "%s", text variable: MAIN_PRG.RobotAction.Planner_ID
        OnMouseClick: write the text variable via Default
    Rectangle (551,660 144x19), "%s", text variable: MAIN_PRG.Status_Error_Codes_Action
    Rectangle (484,363 49x19), "rot_A (Z)"
    Rectangle (484,386 49x19), "rot_B (Y)"
    Rectangle (484,410 49x19), "rot_C (Z)"
    Rectangle (538,364 69x19), "%.3f °", text variable: GVL_OPCUA.rot_A
        OnMouseClick: write the text variable via Default
    Rectangle (538,387 69x19), "%.3f °", text variable: GVL_OPCUA.rot_B
        OnMouseClick: write the text variable via Default
    Rectangle (538,411 69x19), "%.3f °", text variable: GVL_OPCUA.rot_C
        OnMouseClick: write the text variable via Default
    Rectangle (391,441 65x19), "%.3f rad", text variable: MAIN_PRG.RobotAction.joint_tolerance
        OnMouseClick: write the text variable via Default
END_VISUALIZATION
